(* IEC 61131-3 sources: daoli-st-library/DL_Process (part 17) *)

(* ---- FC_DL_RoRecoveryCalc.st ---- *)
(*
  Name: FC_DL_RoRecoveryCalc
  Category: DL_Process
  Version: 1.0.0
  Round: R90 / 2026-11-25
  开源溯源：clean-room 自研（族 RO/NF 膜法水处理，ST 开源生态实测 0 命中，无外部代码引入）
  功能：1) 系统回收率按「产水占进水的百分比」计算，产水为分子、进水为分母，方向固定不可交换，
           即 fRecoveryPct = fPermeateFlowM3h / fFeedFlowM3h * 100，用于 RO/NF 段回收率监视。
        2) 浓水排放流量由容积守恒的减法式给出：进水 − 产水（同温同压下的容积近似），
           作为浓水调节阀的前馈目标值使用。
        3) 回收率同时受两个独立门限约束：物理域 0.0 ~ 100.0 %，以及设计上限
           fRecoveryMaxPct（膜厂家给定的段回收率上限）；任一越界只置 xValid=FALSE，
           数值本身钳制到物理域内后输出，绝不把越限值伪装成合格值。
  边界条件：1) 分母零闸：ABS(fFeedFlowM3h) > DL_EPS 才允许做除法，否则清零全部输出并置无效。
        2) 非有限值闸：全部实值入参先过 NOT(x > -DL_BIG AND x < DL_BIG)，该式同时拦 NaN 与 Inf，
           命中即拦断实值通路（输出强制 0.0），不得只置标志而把 NaN 传给下游（R19）。
        3) 回收率物理域 0.0 ~ 100.0 %，越域钳制到域内输出并置 xValid=FALSE。
        4) 设计上限 fRecoveryMaxPct 自身须落在 (0.0, 100.0] 内，越域视为组态错误判无效。
        5) 产水量为负值（传感器反向）或大于进水量（超出守恒），均判无效，不取绝对值掩盖故障。
        6) 无回差环节：本件为纯函数无状态，不做迟滞，迟滞由下游报警件承担。
  量纲自证：fRecoveryPct = (m3/h) / (m3/h) * 100 = 无因次百分数 [%]；
           fBrineFlowM3h = (m3/h) − (m3/h) = (m3/h)，减法两侧同量纲，量纲关系合法。
*)

FUNCTION FC_DL_RoRecoveryCalc : BOOL
VAR_INPUT
    fFeedFlowM3h     : REAL;   // 系统进水体积流量 [m3/h] / Feed volumetric flow [m3/h]
    fPermeateFlowM3h : REAL;   // 系统产水体积流量 [m3/h] / Permeate volumetric flow [m3/h]
    fRecoveryMaxPct  : REAL;   // 段回收率设计上限 [%] / Design recovery upper limit [%]
END_VAR
VAR_OUTPUT
    fRecoveryPct     : REAL;   // 系统回收率 [%] / System recovery ratio [%]
    fBrineFlowM3h    : REAL;   // 浓水排放流量 [m3/h] / Brine discharge flow [m3/h]
    xValid           : BOOL;   // 计算有效标志 [bool] / Calculation valid flag [bool]
END_VAR
VAR
    _fRecRawPct      : REAL;   // 钳制前的原始回收率 [%] / Raw recovery before limiting [%]
    _fBrineRawM3h    : REAL;   // 钳制前的原始浓水流量 [m3/h] / Raw brine flow before limiting [m3/h]
END_VAR
VAR CONSTANT
    DL_EPS           : REAL := 1.0E-9;    // 分母零闸阈值 [-] / Division-zero gate threshold [-]
    DL_BIG           : REAL := 1.0E12;    // 非有限值闸量级上限 [-] / Finiteness gate magnitude [-]
    DL_PCT           : REAL := 100.0;     // 百分比换算因子 [%] / Percent conversion factor [%]
    DL_REC_LO_PCT    : REAL := 0.0;       // 回收率物理域下限 [%] / Recovery physical domain low [%]
    DL_REC_HI_PCT    : REAL := 100.0;     // 回收率物理域上限 [%] / Recovery physical domain high [%]
END_VAR

(* —— 段 1：非有限值闸（R19：闸断实值通路，NaN/Inf 一律不得流到输出） —— *)
IF NOT (fFeedFlowM3h > -DL_BIG AND fFeedFlowM3h < DL_BIG)
   OR NOT (fPermeateFlowM3h > -DL_BIG AND fPermeateFlowM3h < DL_BIG)
   OR NOT (fRecoveryMaxPct > -DL_BIG AND fRecoveryMaxPct < DL_BIG) THEN
    fRecoveryPct := 0.0;                    // 输出强制 0.0，切断污染源 / Force zero, cut polluted path
    fBrineFlowM3h := 0.0;                   // 浓水同样强制 0.0 / Brine forced to zero as well
    xValid := FALSE;                        // 有效位清零 / Validity cleared
    FC_DL_RoRecoveryCalc := FALSE;          // 返回码与有效位同源 / Return mirrors validity
    RETURN;                                 // 立即退出 / Immediate exit
END_IF

(* —— 段 2：分母零闸（R4：除法前先过 ABS 闸，且闸的是分母本身） —— *)
IF ABS(fFeedFlowM3h) <= DL_EPS THEN
    fRecoveryPct := 0.0;                    // 无进水即无回收率 / No feed means no recovery
    fBrineFlowM3h := 0.0;                   // 无进水即无浓水 / No feed means no brine
    xValid := FALSE;                        // 判无效 / Invalid
    FC_DL_RoRecoveryCalc := FALSE;          // 返回码同步 / Return synchronised
    RETURN;                                 // 提前退出，不做无意义运算 / Early exit
END_IF

(* —— 段 3：主算式（R22 方向自核：差值/比值的基准量是进水量，不是产水量） —— *)
_fRecRawPct := fPermeateFlowM3h / fFeedFlowM3h * DL_PCT;   // 产水 / 进水 * 100 [%]
_fBrineRawM3h := fFeedFlowM3h - fPermeateFlowM3h;          // 进水 − 产水 [m3/h]

(* —— 段 4：物理域与设计上限校验（单点 BOOL 聚合，避免多处赋 FALSE 造成覆盖） —— *)
xValid := (_fRecRawPct >= DL_REC_LO_PCT)                       // 不低于物理域下限
          AND (_fRecRawPct <= DL_REC_HI_PCT)                   // 不高于物理域上限
          AND (fRecoveryMaxPct > DL_EPS)                       // 设计上限必须为正
          AND (fRecoveryMaxPct <= DL_REC_HI_PCT)               // 设计上限不得超 100 %
          AND (_fRecRawPct <= fRecoveryMaxPct)                 // 不得超出膜厂家设计上限
          AND (fPermeateFlowM3h >= 0.0)                        // 产水不得为负（传感器反向）
          AND (fPermeateFlowM3h <= fFeedFlowM3h)               // 产水不得大于进水（守恒校验）
          AND (_fBrineRawM3h >= 0.0);                          // 浓水不得为负

(* —— 段 5：输出单点写盘（数值钳制到物理域内，有效位已在段 4 定案） —— *)
fRecoveryPct := LIMIT(DL_REC_LO_PCT, _fRecRawPct, DL_REC_HI_PCT);   // 回收率钳 0..100 [%]
fBrineFlowM3h := MAX(DL_REC_LO_PCT, _fBrineRawM3h);                 // 浓水钳 >= 0 [m3/h]
FC_DL_RoRecoveryCalc := xValid;                                     // 返回码：TRUE = 计算可信

END_FUNCTION

(* ---- FC_DL_RoScaleSaturationIndexCalc.st ---- *)
(*
  Name: FC_DL_RoScaleSaturationIndexCalc
  Category: DL_Process
  Version: 1.0.0
  Round: R90 / 2026-11-25
  开源溯源：clean-room 自研（族 RO/NF 膜法水处理，ST 开源生态实测 0 命中，无外部代码引入）
  功能：1) 朗格利尔饱和指数按经典四因子式解算：LSI = pH − pHs，
           其中 pHs = (9.3 + A + B) − (C + D)：
             A = (LOG10(TDS) − 1) / 10，表征溶解固体的离子强度；
             B = −13.12 · LOG10(T_K) + 34.55，温度项（T_K 为开尔文，必须做 °C→K 偏移）；
             C = LOG10(Ca 硬度) − 0.4，钙硬度项；
             D = LOG10(碱度)，碱度项。
        2) LOG10 用跨平台安全写法 LN(x) / LN(10) 实现，不依赖厂商私有 LOG10 扩展。
        3) 输出结垢风险等级整数 iRiskLvl：0 = 不结垢（偏腐蚀），1 = 轻度结垢，
           2 = 中度结垢，3 = 严重结垢；等级由 LSI 阈值判定，供加药/阻垢剂投加策略直接取用。
  边界条件：1) 非有限值闸：五路实值入参统一过 NOT(x > -DL_BIG AND x < DL_BIG)，
           同时拦 NaN 与 Inf，命中即拦断实值通路（fLsi 强制 0.0、iRiskLvl 置 0）并置无效（R19）。
        2) 对数自变量零闸：TDS / 钙硬度 / 碱度三项都必须 ABS(x) > DL_EPS 才可进 LN，
           否则 LOG10 发散；任一项不满足判无效。
        3) 对数自变量负值闸：三量均为浓度，负值属变送器故障，判无效且不取 ABS 掩盖。
        4) 量程钳制：TDS 钳 0..60000 mg/L、钙硬度与碱度钳 0..DL_HARD_MAX(2000 mg/L)、
           pH 钳 0..14、温度钳 0..90 °C；越域钳边界值参与计算但置无效。
        5) LSI 结果饱和钳到 −5.0 ~ +5.0 的工程可观测域，防极端输入把指数推到无意义量级。
        6) 无回差环节：纯函数无状态，等级切换的迟滞由下游报警件承担。
  量纲自证：A = (LOG10(mg/L) − 1) / 10 → 无因次 [-]，LOG10 的自变量已按 mg/L 归一；
           B = −13.12 · LOG10(K) + 34.55 → 无因次 [-]，34.55 为经验截距，无单位；
           C、D 同 A 均为无因次；LSI = pH(−) − pHs(−) = 无因次指数 [-]，四项量纲一致。
*)

FUNCTION FC_DL_RoScaleSaturationIndexCalc : BOOL
VAR_INPUT
    fPh              : REAL;   // 给水 pH 值 [pH 单位] / Feed water pH [pH unit]
    fTempC           : REAL;   // 给水温度 [°C] / Feed water temperature [°C]
    fCaHardnessMgL   : REAL;   // 钙硬度（以 CaCO3 计）[mg/L] / Calcium hardness as CaCO3 [mg/L]
    fAlkalinityMgL   : REAL;   // 总碱度（以 CaCO3 计）[mg/L] / Total alkalinity as CaCO3 [mg/L]
    fTdsMgL          : REAL;   // 总溶解固体 [mg/L] / Total dissolved solids [mg/L]
END_VAR
VAR_OUTPUT
    fLsi             : REAL;   // 朗格利尔饱和指数 [-] / Langelier saturation index [-]
    iRiskLvl         : INT;    // 结垢风险等级 0..3 [-] / Scaling risk level 0..3 [-]
    xValid           : BOOL;   // 计算有效标志 [bool] / Calculation valid flag [bool]
END_VAR
VAR
    _fPhClamp        : REAL;   // 钳制后的 pH [-] / Clamped pH [-]
    _fTClampC        : REAL;   // 钳制后的温度 [°C] / Clamped temperature [°C]
    _fCaClampMgL     : REAL;   // 钳制后的钙硬度 [mg/L] / Clamped calcium hardness [mg/L]
    _fAlkClampMgL    : REAL;   // 钳制后的碱度 [mg/L] / Clamped alkalinity [mg/L]
    _fTdsClampMgL    : REAL;   // 钳制后的 TDS [mg/L] / Clamped TDS [mg/L]
    _fTermA          : REAL;   // A 项（TDS 项）[-] / Term A, TDS term [-]
    _fTermB          : REAL;   // B 项（温度项）[-] / Term B, temperature term [-]
    _fTermC          : REAL;   // C 项（钙硬度项）[-] / Term C, calcium hardness term [-]
    _fTermD          : REAL;   // D 项（碱度项）[-] / Term D, alkalinity term [-]
    _fPhs            : REAL;   // 饱和 pH [-] / Saturation pH [-]
    _fLsiRaw         : REAL;   // 未饱和的原始 LSI [-] / Raw LSI before limiting [-]
    _bLogOk          : BOOL;   // 对数自变量合法性聚合 [-] / Logarithm argument validity aggregate
END_VAR
VAR CONSTANT
    DL_EPS           : REAL := 1.0E-9;    // 对数自变量零闸阈值 [-] / Logarithm argument zero gate [-]
    DL_BIG           : REAL := 1.0E12;    // 非有限值闸量级上限 [-] / Finiteness gate magnitude [-]
    DL_K0            : REAL := 273.15;    // 摄氏转开尔文偏移 [K] / Celsius to Kelvin offset [K]
    DL_LN10          : REAL := 2.302585093;   // LN(10)，用于实现 LOG10 [-] / LN(10) for LOG10 [-]
    DL_PH_MAX        : REAL := 14.0;      // pH 量程上限 [-] / pH range high [-]
    DL_T_HI_C        : REAL := 90.0;      // 温度量程上限 [°C] / Temperature range high [°C]
    DL_HARD_MAX      : REAL := 2000.0;    // 钙硬度/碱度量程上限 [mg/L] / Hardness range high [mg/L]
    DL_TDS_MAX       : REAL := 60000.0;   // TDS 量程上限 [mg/L] / TDS range high [mg/L]
    DL_LSI_LO        : REAL := -5.0;      // LSI 工程可观测下限 [-] / LSI observable low [-]
    DL_LSI_HI        : REAL := 5.0;       // LSI 工程可观测上限 [-] / LSI observable high [-]
    DL_LSI_L1        : REAL := 0.0;       // 等级 0/1 分界 [-] / Risk level 0-to-1 boundary [-]
    DL_LSI_L2        : REAL := 0.5;       // 等级 1/2 分界 [-] / Risk level 1-to-2 boundary [-]
    DL_LSI_L3        : REAL := 1.5;       // 等级 2/3 分界 [-] / Risk level 2-to-3 boundary [-]
END_VAR

(* —— 段 1：非有限值闸（R19：五路入参全覆盖，拦 NaN 与 Inf） —— *)
IF NOT (fPh > -DL_BIG AND fPh < DL_BIG)
   OR NOT (fTempC > -DL_BIG AND fTempC < DL_BIG)
   OR NOT (fCaHardnessMgL > -DL_BIG AND fCaHardnessMgL < DL_BIG)
   OR NOT (fAlkalinityMgL > -DL_BIG AND fAlkalinityMgL < DL_BIG)
   OR NOT (fTdsMgL > -DL_BIG AND fTdsMgL < DL_BIG) THEN
    fLsi := 0.0;                            // 输出强制 0.0 / Output forced to zero
    iRiskLvl := 0;                          // 等级置 0（不结垢），不给误导性等级 / Risk level cleared
    xValid := FALSE;                        // 有效位清零 / Validity cleared
    FC_DL_RoScaleSaturationIndexCalc := FALSE;   // 返回码同源 / Return mirrors validity
    RETURN;                                 // 立即退出 / Immediate exit
END_IF

(* —— 段 2：对数自变量零闸 + 负值闸（R4：LN 的自变量必须先验正） —— *)
_bLogOk := (fTdsMgL > DL_EPS) AND (fCaHardnessMgL > DL_EPS) AND (fAlkalinityMgL > DL_EPS);
IF NOT _bLogOk THEN
    fLsi := 0.0;                            // 输出强制 0.0 / Output forced to zero
    iRiskLvl := 0;                          // 等级置 0 / Risk level cleared
    xValid := FALSE;                        // 判无效 / Invalid
    FC_DL_RoScaleSaturationIndexCalc := FALSE;   // 返回码同步 / Return synchronised
    RETURN;                                 // 提前退出 / Early exit
END_IF

(* —— 段 3：量程钳制（边界值参与计算，越域在段 5 判无效） —— *)
_fPhClamp := LIMIT(0.0, fPh, DL_PH_MAX);                  // pH 钳 0..14 [-]
_fTClampC := LIMIT(0.0, fTempC, DL_T_HI_C);               // 温度钳 0..90 [°C]
_fCaClampMgL := LIMIT(0.0, fCaHardnessMgL, DL_HARD_MAX);  // 钙硬度钳 [mg/L]
_fAlkClampMgL := LIMIT(0.0, fAlkalinityMgL, DL_HARD_MAX); // 碱度钳 [mg/L]
_fTdsClampMgL := LIMIT(0.0, fTdsMgL, DL_TDS_MAX);         // TDS 钳 [mg/L]

(* —— 段 4：四因子解算（LOG10 以 LN(x)/LN(10) 跨平台实现） —— *)
_fTermA := (LN(_fTdsClampMgL) / DL_LN10 - 1.0) / 10.0;                          // A 项 [-]
_fTermB := -13.12 * (LN(_fTClampC + DL_K0) / DL_LN10) + 34.55;                  // B 项 [-]
_fTermC := LN(_fCaClampMgL) / DL_LN10 - 0.4;                                    // C 项 [-]
_fTermD := LN(_fAlkClampMgL) / DL_LN10;                                         // D 项 [-]
_fPhs := (9.3 + _fTermA + _fTermB) - (_fTermC + _fTermD);                       // 饱和 pH [-]
_fLsiRaw := _fPhClamp - _fPhs;                                                  // LSI = pH − pHs [-]

(* —— 段 5：有效位单点聚合（量程校验，钳制值已参与计算） —— *)
xValid := (fPh >= 0.0) AND (fPh <= DL_PH_MAX)                                   // pH 在量程内
          AND (fTempC >= 0.0) AND (fTempC <= DL_T_HI_C)                         // 温度在量程内
          AND (fCaHardnessMgL <= DL_HARD_MAX)                                   // 钙硬度不越上限
          AND (fAlkalinityMgL <= DL_HARD_MAX)                                   // 碱度不越上限
          AND (fTdsMgL <= DL_TDS_MAX);                                          // TDS 不越上限

(* —— 段 6：风险等级分级（IF/ELSIF 单链，iRiskLvl 只在此处赋值一次） —— *)
IF _fLsiRaw < DL_LSI_L1 THEN
    iRiskLvl := 0;                          // 不结垢（偏腐蚀倾向）/ Non-scaling, corrosive tendency
ELSIF _fLsiRaw < DL_LSI_L2 THEN
    iRiskLvl := 1;                          // 轻度结垢 / Slight scaling tendency
ELSIF _fLsiRaw < DL_LSI_L3 THEN
    iRiskLvl := 2;                          // 中度结垢 / Moderate scaling tendency
ELSE
    iRiskLvl := 3;                          // 严重结垢 / Severe scaling tendency
END_IF

(* —— 段 7：输出单点写盘（LSI 饱和钳到工程可观测域） —— *)
fLsi := LIMIT(DL_LSI_LO, _fLsiRaw, DL_LSI_HI);   // LSI 钳 −5..+5 [-]
FC_DL_RoScaleSaturationIndexCalc := xValid;      // 返回码：TRUE = 计算可信

END_FUNCTION

(* ---- FC_DL_RoStagePressureDropCalc.st ---- *)
(*
  Name: FC_DL_RoStagePressureDropCalc
  Category: DL_Process
  Version: 1.0.0
  Round: R90 / 2026-11-25
  开源溯源：clean-room 自研（族 RO/NF 膜法水处理，ST 开源生态实测 0 命中，无外部代码引入）
  功能：1) 段间压降按湍流平方律计算：ΔP = k · Q²，其中 k 为段阻力系数（bar/(m3/h)²），
           Q 为段流量（m3/h）。平方律的依据是湍流区沿程与局部损失均与流速平方成正比，
           而流速与容积流量成正比，故压降对流量呈二次关系，不是线性关系。
        2) 与压降上限 fDropLimitBar 比对给出超限报警 xAlarm。超限是膜段污堵/浓水通道阻塞的
           早期特征（流量不变而压降上升），因此报警取「大于等于上限」而非「大于」，
           上限触点本身即算到达报警点。
  边界条件：1) 非有限值闸：三路实值入参统一过 NOT(x > -DL_BIG AND x < DL_BIG)，
           同时拦 NaN 与 Inf，命中即拦断实值通路（fDropBar 强制 0.0、xAlarm 强制 FALSE）并置无效（R19）。
        2) 组态零闸：ABS(fResistCoef) > DL_EPS 与 ABS(fDropLimitBar) > DL_EPS 都必须成立，
           阻力系数为 0 表示未标定、上限为 0 表示未组态，两者都判无效（不做除零以外的默认替代）。
        3) 负值闸：段流量为负判无效（传感器反向）；阻力系数为负判无效（系数不可为负）；
           压降上限为负判无效。
        4) 饱和钳制：段流量先钳到 0 ~ DL_FLOW_MAX(1000 m3/h)，压降结果再钳到 0 ~ DL_DROP_MAX(50 bar)，
           防止平方项在小数域溢出或给出无物理意义的巨值。
        5) 报警只在 xValid 为 TRUE 时才可能为 TRUE，无效数据不得触发工艺报警（防误停）。
        6) 无回差环节：本件为纯函数无状态，报警回差由下游 FB 承担。
  量纲自证：ΔP = (bar/(m3/h)²) × (m3/h)² = bar，平方项与系数分母量纲对消，量纲闭合；
           报警比较两侧同为 bar，量纲一致，禁止与 kPa 混比。
*)

FUNCTION FC_DL_RoStagePressureDropCalc : BOOL
VAR_INPUT
    fStageFlowM3h    : REAL;   // 段内体积流量 [m3/h] / Stage volumetric flow [m3/h]
    fResistCoef      : REAL;   // 段阻力系数 [bar/(m3/h)²] / Stage resistance coefficient [bar/(m3/h)^2]
    fDropLimitBar    : REAL;   // 段间压降报警上限 [bar] / Pressure drop alarm limit [bar]
END_VAR
VAR_OUTPUT
    fDropBar         : REAL;   // 段间压降 [bar] / Stage pressure drop [bar]
    xAlarm           : BOOL;   // 压降超限报警 [bool] / Pressure drop over-limit alarm [bool]
    xValid           : BOOL;   // 计算有效标志 [bool] / Calculation valid flag [bool]
END_VAR
VAR
    _fFlowClampM3h   : REAL;   // 钳制后的段流量 [m3/h] / Clamped stage flow [m3/h]
    _fDropRawBar     : REAL;   // 未饱和的原始压降 [bar] / Raw pressure drop [bar]
END_VAR
VAR CONSTANT
    DL_EPS           : REAL := 1.0E-9;    // 组态零闸阈值 [-] / Configuration zero gate threshold [-]
    DL_BIG           : REAL := 1.0E12;    // 非有限值闸量级上限 [-] / Finiteness gate magnitude [-]
    DL_FLOW_MAX      : REAL := 1000.0;    // 段流量饱和钳制上限 [m3/h] / Stage flow saturation ceiling [m3/h]
    DL_DROP_MAX      : REAL := 50.0;      // 压降饱和钳制上限 [bar] / Pressure drop saturation ceiling [bar]
END_VAR

(* —— 段 1：非有限值闸（R19：三路入参全覆盖，拦 NaN 与 Inf） —— *)
IF NOT (fStageFlowM3h > -DL_BIG AND fStageFlowM3h < DL_BIG)
   OR NOT (fResistCoef > -DL_BIG AND fResistCoef < DL_BIG)
   OR NOT (fDropLimitBar > -DL_BIG AND fDropLimitBar < DL_BIG) THEN
    fDropBar := 0.0;                        // 输出强制 0.0 / Output forced to zero
    xAlarm := FALSE;                        // 报警强制 FALSE，无效数据不得触发停运 / Alarm forced off
    xValid := FALSE;                        // 有效位清零 / Validity cleared
    FC_DL_RoStagePressureDropCalc := FALSE; // 返回码同源 / Return mirrors validity
    RETURN;                                 // 立即退出 / Immediate exit
END_IF

(* —— 段 2：组态零闸（阻力系数与报警上限都必须已标定，0 值视为未组态） —— *)
IF (ABS(fResistCoef) <= DL_EPS) OR (ABS(fDropLimitBar) <= DL_EPS) THEN
    fDropBar := 0.0;                        // 输出强制 0.0 / Output forced to zero
    xAlarm := FALSE;                        // 报警强制 FALSE / Alarm forced off
    xValid := FALSE;                        // 判无效 / Invalid
    FC_DL_RoStagePressureDropCalc := FALSE; // 返回码同步 / Return synchronised
    RETURN;                                 // 提前退出 / Early exit
END_IF

(* —— 段 3：负值闸（流量反向 / 系数为负 / 上限为负，三者均属组态或传感器故障） —— *)
IF (fStageFlowM3h < 0.0) OR (fResistCoef < 0.0) OR (fDropLimitBar < 0.0) THEN
    fDropBar := 0.0;                        // 输出强制 0.0 / Output forced to zero
    xAlarm := FALSE;                        // 报警强制 FALSE / Alarm forced off
    xValid := FALSE;                        // 判无效 / Invalid
    FC_DL_RoStagePressureDropCalc := FALSE; // 返回码同步 / Return synchronised
    RETURN;                                 // 提前退出 / Early exit
END_IF

(* —— 段 4：平方律主算式（R22 方向自核：流量平方乘系数，非系数除流量） —— *)
_fFlowClampM3h := LIMIT(0.0, fStageFlowM3h, DL_FLOW_MAX);    // 流量钳 0..1000 [m3/h]
_fDropRawBar := fResistCoef * _fFlowClampM3h * _fFlowClampM3h;   // ΔP = k·Q² [bar]

(* —— 段 5：输出单点写盘（先饱和钳制，再据此判报警，保证判据用的是同一个值） —— *)
fDropBar := LIMIT(0.0, _fDropRawBar, DL_DROP_MAX);           // 压降钳 0..50 [bar]
xValid := (fResistCoef > DL_EPS)                             // 系数已标定且为正
          AND (fDropLimitBar > DL_EPS)                       // 上限已组态且为正
          AND (fStageFlowM3h >= 0.0);                        // 流量非负
xAlarm := xValid AND (fDropBar >= fDropLimitBar);            // 到达上限即报警（含触点）

(* —— 段 6：返回码（TRUE = 计算可信，与 xValid 同源） —— *)
FC_DL_RoStagePressureDropCalc := xValid;

END_FUNCTION

(* ---- FC_DL_SandToMetalRatioCalc.st ---- *)
(*
 * FC_DL_SandToMetalRatioCalc | C1 | DL_Process
 * 功能：砂铁比（单位铸铁合格件对应的砂循环量）       单位：流量 [kg/h]、比值 [kg/kg]
 * 工况边界：仅适用于连续生产的砂处理线（砂循环量与铁水消耗量同口径统计）；金属流量须 >0（入分母），砂流量须 ≥0 且有限；不区分新旧砂，只算总量比值
 * 代数值回代：sand=120000 kg/h、metal=15000 kg/h → 比值 8.0 kg/kg（与 spec 回代行一致）
 * 开源溯源：clean-room 自研，未复制任何第三方代码（无外部来源）
 *)
FUNCTION FC_DL_SandToMetalRatioCalc : BOOL
VAR_INPUT
    rSandKgH  : REAL := 120000.0;    // 砂循环量 | sand circulation rate [kg/h]
    rMetalKgH : REAL := 15000.0;     // 铁水消耗量 | molten metal consumption rate [kg/h]
END_VAR
VAR_OUTPUT
    rRatio     : REAL;               // 砂铁比 | sand to metal ratio [kg/kg]
    xValid     : BOOL;               // 输出有效 | outputs valid
    nFaultCode : INT;                // 0=无 / 9711=金属流量非法 | 0 none, 9711 illegal metal flow
END_VAR
VAR
    xFinSand  : BOOL;                // 砂流量有限性 | sand flow is finite
    xFinMetal : BOOL;                // 金属流量有限性 | metal flow is finite
END_VAR
VAR CONSTANT
    DL_SMR_METAL_MIN : REAL := 1.0E-9;  // 金属流量下限（防零除）| metal flow lower bound [kg/h]
END_VAR

// 段1｜非有限闸（R19）
xFinSand := (rSandKgH = rSandKgH) AND ((rSandKgH - rSandKgH) = 0.0);
xFinMetal := (rMetalKgH = rMetalKgH) AND ((rMetalKgH - rMetalKgH) = 0.0);
IF (NOT xFinSand) OR (NOT xFinMetal) THEN
    rRatio := 0.0;                   // 安全值：比值 0 | safe value, zero ratio
    xValid := FALSE;
    nFaultCode := 9711;
    FC_DL_SandToMetalRatioCalc := FALSE;
    RETURN;
END_IF

// 段2｜域闸：金属流量入分母必须 >0，砂流量不得为负
IF (rMetalKgH <= DL_SMR_METAL_MIN) OR (rSandKgH < 0.0) THEN
    rRatio := 0.0;
    xValid := FALSE;
    nFaultCode := 9711;
    FC_DL_SandToMetalRatioCalc := FALSE;
    RETURN;
END_IF

// 段3｜算法与出口
rRatio := rSandKgH / rMetalKgH;
nFaultCode := 0;
xValid := TRUE;
FC_DL_SandToMetalRatioCalc := TRUE;
END_FUNCTION

(* ---- FC_DL_SanitizeHoldTimeCalc.st ---- *)
(*
  ============================================================
  组件名 : FC_DL_SanitizeHoldTimeCalc
  分类   : DL_Process
  功能   : 消毒保持时间计算，按实际浓度折算浓度比并对温度系数修正后给出保持时间
  复杂度 : C1
  版本   : 1.0.0
  作者   : 道莅工业代码库工厂 / R81
  日期   : 2026-11-24
  开源溯源 : clean-room（no upstream）—— 依据公开工程公式自研，未复制任何上游实现
  红线自检 : R1 无GVL/R2 无物理地址/R3 纯IEC/R4 防除零/R5 双语注释
  接口说明 :
      温度系数 = 1 + (温度-20)*0.02，限幅 0.5~2.0，防止极端温度把时间推到无意义区间。
      保持时间 = 基准时间 * (基准浓度/实际浓度) * (1/温度系数)。
      浓度低于基准时比值大于 1，时间自动延长；浓度高于基准时时间缩短，符合消毒动力学方向。
  ============================================================
*)
FUNCTION FC_DL_SanitizeHoldTimeCalc : BOOL
VAR_INPUT
    bEnable      : BOOL; // 使能：TRUE 时计算 / Enable: TRUE to compute
    bErr         : BOOL; // 外部故障：TRUE 时立即退出并置结果无效 / External fault: TRUE aborts with invalid result
    rConcPct     : REAL; // 实际消毒液浓度 [%] / actual sanitizer concentration [percent]
    rConcRefPct  : REAL; // 基准消毒液浓度 [%] / reference sanitizer concentration [percent]
    rHoldRef_min : REAL; // 基准浓度下的基准保持时间 [min] / reference hold time at the reference concentration [minute]
    rTempC       : REAL; // 实际消毒液温度 [摄氏度] / actual sanitizer temperature [degree Celsius]
END_VAR
VAR_OUTPUT
    rTempFactor : REAL; // 温度修正系数，限幅 0.5~2.0 [无量纲] / temperature correction factor clamped to 0.5 to 2.0 [dimensionless]
    rConcRatio  : REAL; // 浓度比，基准浓度除以实际浓度 [无量纲] / concentration ratio of reference over actual [dimensionless]
    rHold_min   : REAL; // 修正后的保持时间 [min] / corrected hold time [minute]
    bValid      : BOOL; // 输出有效：TRUE 表示结果可用 / Output valid
END_VAR
VAR CONSTANT
    DL_R_MAX    : REAL := 3.0E38; // 实数上界，用于拦截 Inf [无量纲] / real upper bound used to reject infinity [dimensionless]
    DL_EPS      : REAL := 1.0E-12; // 除零判定阈值 [无量纲] / division guard threshold [dimensionless]
    DL_ONE      : REAL := 1.0;    // 单位常量 [无量纲] / unity constant [dimensionless]
    DL_TEMP_REF : REAL := 20.0;   // 温度基准点 [摄氏度] / temperature reference point [degree Celsius]
    DL_TEMP_K   : REAL := 0.02;   // 每摄氏度温度系数增量 [1/摄氏度] / temperature coefficient increment per degree Celsius [per degree Celsius]
    DL_FACT_LO  : REAL := 0.5;    // 温度系数下限 [无量纲] / lower limit of the temperature factor [dimensionless]
    DL_FACT_HI  : REAL := 2.0;    // 温度系数上限 [无量纲] / upper limit of the temperature factor [dimensionless]
    DL_TEMP_MIN : REAL := -50.0;  // 允许温度下界 [摄氏度] / permitted lower bound of the temperature [degree Celsius]
    DL_TEMP_MAX : REAL := 150.0;  // 允许温度上界 [摄氏度] / permitted upper bound of the temperature [degree Celsius]
END_VAR
VAR
    _bFin  : BOOL := FALSE; // 输入有限性判定结果 / input finiteness verdict
    _rInv  : REAL := 0.0;   // 温度系数的倒数，除法前先算后判 [无量纲] / reciprocal of the temperature factor computed before the guard [dimensionless]
END_VAR

    // 段 1｜出口预置：系数先置于 1，避免下游误用零
    rTempFactor := DL_ONE;
    rConcRatio := 0.0;
    rHold_min := 0.0;
    bValid := FALSE;
    // 段 2｜使能闸与外部故障闸
    IF NOT bEnable THEN
        RETURN;
    END_IF;
    IF bErr THEN
        RETURN;
    END_IF;
    // 段 3｜非有限闸
    _bFin := (rConcPct = rConcPct) AND (ABS(rConcPct) <= DL_R_MAX) AND (rConcRefPct = rConcRefPct) AND (ABS(rConcRefPct) <= DL_R_MAX) AND (rHoldRef_min = rHoldRef_min) AND (ABS(rHoldRef_min) <= DL_R_MAX) AND (rTempC = rTempC) AND (ABS(rTempC) <= DL_R_MAX);
    IF NOT _bFin THEN
        RETURN;
    END_IF;
    // 段 4｜域闸：实际浓度严格为正、基准浓度非负、基准时间非负、温度在工程区间
    IF ABS(rConcPct) <= DL_EPS THEN
        RETURN;
    END_IF;
    IF (rConcPct < 0.0) OR (rConcRefPct < 0.0) OR (rHoldRef_min < 0.0) THEN
        RETURN;
    END_IF;
    IF (rTempC < DL_TEMP_MIN) OR (rTempC > DL_TEMP_MAX) THEN
        RETURN;
    END_IF;
    // 段 5｜温度系数与限幅
    rTempFactor := DL_ONE + (rTempC - DL_TEMP_REF) * DL_TEMP_K;
    IF rTempFactor > DL_FACT_HI THEN
        rTempFactor := DL_FACT_HI;
    ELSIF rTempFactor < DL_FACT_LO THEN
        rTempFactor := DL_FACT_LO;
    END_IF;
    // 段 6｜浓度比
    rConcRatio := rConcRefPct / rConcPct;
    // 段 7｜温度系数分母闸：先判零再取倒数，顺序不可颠倒
    IF ABS(rTempFactor) <= DL_EPS THEN
        RETURN;
    END_IF;
    _rInv := DL_ONE / rTempFactor;
    rHold_min := rHoldRef_min * rConcRatio * _rInv;
    bValid := TRUE;
    FC_DL_SanitizeHoldTimeCalc := bValid;
END_FUNCTION

(* ---- FC_DL_ScreenEfficiencyCalc.st ---- *)
(*
  Name: FC_DL_ScreenEfficiencyCalc
  Category: DL_Process
  Version: 1.0.0
  Round: R89 / 2026-11-25
  开源溯源：clean-room 自研（族 矿山破碎筛分，ST 开源生态实测 0 命中，无外部代码引入）
  功能：按入料/筛上/筛下三处细粒含量算振动筛筛分效率（经典式，全部折算为小数参与运算）。
  边界条件：① 三入参百分数先折算小数，入料细粒 0~100 %、筛上 0~100 %、筛下 0~100 %；
            ② 分母 (1−O)·(F+U−1) 显式零闸，绝对值不超 DL_EPS 即判非法返回哨兵 -1；
            ③ 效率物理域 0~100 %；算得负值（物料衡算矛盾，如筛下含量低于入料）判 xValid = FALSE 并返回 -1。
  量纲自证：F/O/U 均为质量分数（无量纲），E 亦无量纲，×100 得百分数。
*)
FUNCTION FC_DL_ScreenEfficiencyCalc : REAL
VAR_INPUT
    fFeedFinesPct : REAL;   (* 入料细粒含量 [%] Feed fines content [%] *)
    fOverFinesPct : REAL;   (* 筛上细粒含量 [%] Oversize fines content [%] *)
    fUnderFinesPct : REAL;  (* 筛下合格细粒含量 [%] Undersize fines content [%] *)
END_VAR
VAR_OUTPUT
    fEfficiencyPct : REAL;  (* 筛分效率 [%] Screening efficiency [%] *)
    xValid : BOOL;          (* 计算有效性标志 [-] Calculation valid flag *)
END_VAR
VAR CONSTANT
    DL_EPS : REAL := 1.0E-9;    (* 除零判定容差 [-] Divide-by-zero tolerance *)
    DL_PCT : REAL := 100.0;     (* 百分数基准 [%] Percent base *)
    DL_E_MAX : REAL := 100.0;   (* 效率饱和上限 [%] Efficiency ceiling *)
END_VAR
VAR
    fF : REAL;      (* 入料细粒质量分数 [-] Feed fines fraction *)
    fO : REAL;      (* 筛上细粒质量分数 [-] Oversize fines fraction *)
    fU : REAL;      (* 筛下细粒质量分数 [-] Undersize fines fraction *)
    fDen : REAL;    (* 分母 (1−O)·(F+U−1) [-] Denominator *)
    fEff : REAL;    (* 效率小数中间量 [-] Efficiency scratch *)
END_VAR
(* 出口预置：两出口统一预置（R256） *)
fEfficiencyPct := 0.0; xValid := FALSE;
(* 非有限闸：NaN 自反判 + Inf 差值自减判，三入参全枚举 *)
IF (fFeedFinesPct <> fFeedFinesPct) OR ((fFeedFinesPct - fFeedFinesPct) <> 0.0)
   OR (fOverFinesPct <> fOverFinesPct) OR ((fOverFinesPct - fOverFinesPct) <> 0.0)
   OR (fUnderFinesPct <> fUnderFinesPct) OR ((fUnderFinesPct - fUnderFinesPct) <> 0.0) THEN
    FC_DL_ScreenEfficiencyCalc := -1.0;     (* 哨兵 -1：入参非有限 / Sentinel -1, non-finite input *)
    RETURN;
END_IF
(* 组态域闸：三处含量皆须落在 0~100 %，入料细粒须 > 0（为除子） *)
IF (fFeedFinesPct <= DL_EPS) OR (fFeedFinesPct > DL_PCT)
   OR (fOverFinesPct < 0.0) OR (fOverFinesPct >= DL_PCT)
   OR (fUnderFinesPct < 0.0) OR (fUnderFinesPct > DL_PCT) THEN
    FC_DL_ScreenEfficiencyCalc := -1.0;     (* 哨兵 -1：组态非法 / Sentinel -1, bad configuration *)
    RETURN;
END_IF
(* 百分数折算小数，量纲变为质量分数 *)
fF := fFeedFinesPct / DL_PCT;
fO := fOverFinesPct / DL_PCT;
fU := fUnderFinesPct / DL_PCT;
(* 经典二产品筛分效率式分母：D = F·(U−O)，先算后闸，禁先除后判 *)
(* 原式 D=(1−O)(F+U−1) 会把 η 放大 1/(F+U−1) 倍并系统性饱和到 100%，已废弃 *)
fDen := fF * (fU - fO);
IF ABS(fDen) <= DL_EPS THEN
    FC_DL_ScreenEfficiencyCalc := -1.0;     (* 哨兵 -1：分母塌零 / Sentinel -1, vanishing denominator *)
    RETURN;
END_IF
(* E = U·(F−O) / (F·(U−O))，F 已过零闸，D 已过塌零闸（Wills 选矿手册式） *)
fEff := (fU * (fF - fO)) / fDen;
(* 负值即物料衡算矛盾（筛下细粒反少于入料平衡），判非法不钳成 0 冒充正常 *)
IF fEff < -DL_EPS THEN
    FC_DL_ScreenEfficiencyCalc := -1.0;     (* 哨兵 -1：衡算矛盾 / Sentinel -1, mass-balance conflict *)
    RETURN;
END_IF
(* 物理域钳位：效率不超 100 %，微负残差按 0 处理 *)
IF fEff > 1.0 THEN
    fEff := 1.0;                            (* 上限钳位 100 % / Clamp to 100 percent *)
ELSIF fEff < 0.0 THEN
    fEff := 0.0;                            (* 微负残差归零 / Negative residual to zero *)
END_IF
fEfficiencyPct := fEff * DL_PCT;            (* 分数 → 百分数 [%] Fraction to percent *)
xValid := TRUE;                             (* 链路有效 / Chain valid *)
FC_DL_ScreenEfficiencyCalc := fEfficiencyPct;
END_FUNCTION

(* ---- FC_DL_ScrewPressThroughput.st ---- *)
(*
  道莅工业代码库 / Daoli Industrial ST Library
  组件: FC_DL_ScrewPressThroughput
  分类: DL_Process
  开源溯源: 无（clean-room 工程公式自研；参考公开工艺计算公式，未复制任何受版权保护代码）
  许可证: 本项目自有 (MIT)
  功能: 螺旋压榨机干固体（DS）处理量换算：小时量与按日运行小时数折算的日总量
*)
FUNCTION FC_DL_ScrewPressThroughput : BOOL
VAR_INPUT
    rFlowM3h : REAL; // 进泥体积流量 [m3/h] / sludge feed flow
    rTsPct : REAL; // 进泥含固率 [%] / feed total solids content
    rRunHours : REAL; // 日运行小时数 [h/d] / daily running hours
END_VAR
VAR_OUTPUT
    rDsKgH : REAL; // 干固体小时处理量 [kg/h] / dry solids throughput per hour
    rDsKgDay : REAL; // 干固体日处理量 [kg/d] / dry solids throughput per day
    bValid : BOOL; // 结果有效位 [-] / result valid flag
    iErrCode : INT; // 事件码 0=正常 1=含固率超域 2=运行小时超域 3=结果非有限 / event code
END_VAR
VAR CONSTANT
    rRhoSludge : REAL := 1000.0; // 污泥近似密度 [kg/m3] / approximate sludge density
    rPctToFrac : REAL := 0.01; // 百分数转小数系数 [-]/[%] / percent to fraction factor
    rHourPerDay : REAL := 24.0; // 每日小时数 [h/d] / hours per day
END_VAR
VAR
    rDsRaw : REAL; // 未校验小时量 [kg/h] / unchecked hourly throughput
END_VAR

    // —— 段 0：全路径预清 —— //
    rDsRaw := 0.0;
    rDsKgH := 0.0;
    rDsKgDay := 0.0;
    bValid := FALSE;
    iErrCode := 0;
    FC_DL_ScrewPressThroughput := FALSE;
    // —— 段 1：含固率域闸 (0, 100]% —— //
    IF (rTsPct <= 0.0) OR (rTsPct > 100.0) THEN
        iErrCode := 1; // 含固率超域，干固体量无意义 / TS out of domain, dry solids meaningless
        RETURN;
    END_IF;
    // —— 段 2：日运行小时域闸 (0, 24]h —— //
    IF (rRunHours <= 0.0) OR (rRunHours > rHourPerDay) THEN
        iErrCode := 2; // 运行小时超域 / running hours out of domain
        RETURN;
    END_IF;
    // —— 段 3：量纲链 (m3/h)*(kg/m3)*(%)*(0.01) = kg/h —— //
    rDsRaw := rFlowM3h * rRhoSludge * rTsPct * rPctToFrac; // 干固体量 [kg/h] / dry solids per hour
    IF ABS(rDsRaw) > 1.0E15 THEN
        iErrCode := 3; // 结果非有限，强制归零 / non-finite result, forced to zero
        RETURN;
    END_IF;
    IF rDsRaw < 0.0 THEN
        rDsKgH := 0.0; // 负流量防御 / negative flow guard
    ELSE
        rDsKgH := rDsRaw;
    END_IF;
    // —— 段 4：日总量 = 小时量 × 日运行小时（量纲 kg/h × h/d = kg/d） —— //
    rDsKgDay := rDsKgH * rRunHours; // 日处理量 [kg/d] / dry solids per day
    bValid := TRUE;
    FC_DL_ScrewPressThroughput := TRUE;
END_FUNCTION

(* ---- FC_DL_ScrubberLiquidGasRatio.st ---- *)
(*
  道莅工业代码库 / Daoli Industrial ST Library
  组件: FC_DL_ScrubberLiquidGasRatio
  分类: DL_Process
  开源溯源: 无（clean-room 工程公式自研；参考公开工艺计算公式，未复制任何受版权保护代码）
  许可证: 本项目自有 (MIT)
  功能: 湿式洗涤塔液气比（L/m3）计算、最低液量需求与低液气比告警
*)
FUNCTION FC_DL_ScrubberLiquidGasRatio : BOOL
VAR_INPUT
    rLiquidM3h : REAL; // 循环液流量 [m3/h] / scrubbing liquid flow
    rGasNm3h : REAL; // 标态烟气量 [Nm3/h] / flue gas flow at normal conditions
END_VAR
VAR_OUTPUT
    rLG : REAL; // 液气比 [L/m3] / liquid to gas ratio
    rLiquidNeedM3h : REAL; // 满足最低液气比所需液量 [m3/h] / liquid demand at the minimum ratio
    bValid : BOOL; // 结果有效位 [-] / result valid flag
    bLow : BOOL; // 低液气比告警（<2.0 L/m3）[-] / low ratio alarm
    iErrCode : INT; // 事件码 0=正常 1=烟气量非法 2=结果非有限 / event code
END_VAR
VAR CONSTANT
    rM3ToL : REAL := 1000.0; // 立方米转升系数 [L/m3] / cubic metre to litre factor
    rLgMin : REAL := 2.0; // 最低液气比 [L/m3] / minimum liquid to gas ratio
END_VAR
VAR
    rLgRaw : REAL; // 未限幅液气比 [L/m3] / unlimited ratio
    rNeedLh : REAL; // 最低液量需求 [L/h] / liquid demand in L/h
END_VAR

    // —— 段 0：全路径预清 —— //
    rLgRaw := 0.0;
    rNeedLh := 0.0;
    rLG := 0.0;
    rLiquidNeedM3h := 0.0;
    bValid := FALSE;
    bLow := FALSE;
    iErrCode := 0;
    FC_DL_ScrubberLiquidGasRatio := FALSE;
    // —— 段 1：分母闸（烟气量必须为正） —— //
    IF rGasNm3h <= 0.0 THEN
        iErrCode := 1; // 烟气量非法，液气比无定义 / invalid gas flow, ratio undefined
        RETURN;
    END_IF;
    // —— 段 2：量纲链 (m3/h)/(Nm3/h) = 无量纲，×(L/m3) 得 L/m3 —— //
    rLgRaw := rLiquidM3h / rGasNm3h * rM3ToL; // 液气比 [L/m3] / liquid to gas ratio
    IF ABS(rLgRaw) > 1.0E15 THEN
        iErrCode := 2; // 结果非有限，强制归零 / non-finite result, forced to zero
        RETURN;
    END_IF;
    IF rLgRaw < 0.0 THEN
        rLG := 0.0; // 负液量防御 / negative liquid guard
    ELSE
        rLG := rLgRaw;
    END_IF;
    // —— 段 3：最低液量反算（量纲 (L/m3)×(Nm3/h)/(L/m3) = m3/h） —— //
    rNeedLh := rLgMin * rGasNm3h; // 最低液量 [L/h] / minimum liquid in L/h
    rLiquidNeedM3h := rNeedLh / rM3ToL; // 折算 m3/h / back to m3/h
    // —— 段 4：低液气比告警（信息级，数值照给） —— //
    bLow := rLG < rLgMin; // 低液气比标志 [-] / low ratio flag
    bValid := TRUE;
    FC_DL_ScrubberLiquidGasRatio := TRUE;
END_FUNCTION

(* ---- FC_DL_SettleVelocityCalc.st ---- *)
(*
  道莅工业代码库 / Daoli Industrial ST Library
  组件: FC_DL_SettleVelocityCalc
  分类: DL_Process
  开源溯源: 无（clean-room 工程公式自研；参考公开工艺计算公式，未复制任何受版权保护代码）
  许可证: 本项目自有 (MIT)
  功能: Stokes 自由沉降末速度，含雷诺数域校验（Re>2 判为超出 Stokes 层流域）
*)
FUNCTION FC_DL_SettleVelocityCalc : BOOL
VAR_INPUT
    rDpUm : REAL; // 颗粒粒径 [µm] / particle diameter in micrometre
    rRhoP : REAL; // 颗粒密度 [kg/m3] / particle density
    rRhoF : REAL; // 流体密度 [kg/m3] / fluid density
    rMuPas : REAL; // 流体动力黏度 [mPa·s] / dynamic viscosity in mPa·s
END_VAR
VAR_OUTPUT
    rVsMmS : REAL; // 沉降末速度 [mm/s] / terminal settling velocity
    bValid : BOOL; // 结果有效位（超出 Stokes 域时置 FALSE）[-] / valid flag, FALSE when outside Stokes regime
    iErrCode : INT; // 事件码 0=正常 1=黏度非法 2=密度差不正（按 0 处理）3=Re 超域 4=结果非有限 / event code
END_VAR
VAR CONSTANT
    rGravity : REAL := 9.80665; // 标准重力加速度 [m/s2] / standard gravity
    rUmToM : REAL := 1.0E-6; // 微米转米系数 [m/µm] / micrometre to metre factor
    rMpasToPas : REAL := 1.0E-3; // 毫帕秒转帕秒系数 [Pa·s/(mPa·s)] / mPa·s to Pa·s factor
    rStokesCoef : REAL := 18.0; // Stokes 阻力式系数（无量纲）[-] / Stokes drag coefficient
    rReLimit : REAL := 2.0; // Stokes 层流域上界雷诺数 [-] / upper Reynolds number of Stokes regime
END_VAR
VAR
    rDm : REAL; // 颗粒粒径 [m] / particle diameter in metre
    rMuPas2 : REAL; // 动力黏度 [Pa·s] / dynamic viscosity in Pa·s
    rVsMs : REAL; // 沉降末速度 [m/s] / terminal velocity in m/s
    rRe : REAL; // 颗粒雷诺数 [-] / particle Reynolds number
END_VAR

    // —— 段 0：全路径预清 —— //
    rDm := 0.0;
    rMuPas2 := 0.0;
    rVsMs := 0.0;
    rRe := 0.0;
    rVsMmS := 0.0;
    bValid := FALSE;
    iErrCode := 0;
    FC_DL_SettleVelocityCalc := FALSE;
    // —— 段 1：分母闸（黏度）与单位归一到 SI —— //
    IF rMuPas <= 0.0 THEN
        iErrCode := 1; // 黏度非正，Stokes 式无定义 / non-positive viscosity, Stokes law undefined
        RETURN;
    END_IF;
    rMuPas2 := rMuPas * rMpasToPas; // [mPa·s] -> [Pa·s] / viscosity to SI
    rDm := rDpUm * rUmToM; // [µm] -> [m] / diameter to SI
    // —— 段 2：不上浮判据（固相密度不大于液相时按零速处理） —— //
    IF rRhoP <= rRhoF THEN
        rVsMmS := 0.0;
        iErrCode := 2; // 密度差不正，颗粒不沉降 / non-positive density difference, no settling
        RETURN;
    END_IF;
    // —— 段 3：量纲链 (m/s2)*(m2)*(kg/m3)/(Pa·s) = m/s —— //
    rVsMs := rGravity * rDm * rDm * (rRhoP - rRhoF) / (rStokesCoef * rMuPas2); // 末速度 [m/s] / terminal velocity
    IF ABS(rVsMs) > 1.0E15 THEN
        rVsMs := 0.0;
        iErrCode := 4; // 结果非有限，强制归零 / non-finite result, forced to zero
        RETURN;
    END_IF;
    // —— 段 4：Re 校验（d*v*rhoF/mu），超 2 即离开 Stokes 层流域 —— //
    rRe := rDm * rVsMs * rRhoF / rMuPas2; // 雷诺数 [-] / particle Reynolds number
    rVsMmS := rVsMs * 1000.0; // [m/s] -> [mm/s] / velocity to mm/s
    IF rRe > rReLimit THEN
        iErrCode := 3; // 超出 Stokes 域，给值但标无效 / outside Stokes regime, value kept but flagged
        bValid := FALSE;
        FC_DL_SettleVelocityCalc := FALSE;
        RETURN;
    END_IF;
    bValid := TRUE;
    FC_DL_SettleVelocityCalc := TRUE;
END_FUNCTION

(* ---- FC_DL_ShadeDriftIndexCalc.st ---- *)
(*
  DL Factory R83 | FC_DL_ShadeDriftIndexCalc
  功能：把 L*a*b* 三通道色差按亮度权重合成为色差与漂移指数，并给出回修判定。
  开源溯源：无（clean-room 自研，依据公开工艺公式，来源=行业通用公式，许可证=MIT，借鉴点=公式结构）
  规则：R1-R21 全遵守
*)
FUNCTION FC_DL_ShadeDriftIndexCalc : REAL
VAR_INPUT
    fDeltaL  : REAL; // 明度差 ΔL（正=偏亮）[ΔE 单位] / Lightness difference [dE]
    fDeltaA  : REAL; // 红绿轴差 Δa（正=偏红）[ΔE 单位] / Red-green difference [dE]
    fDeltaB  : REAL; // 黄蓝轴差 Δb（正=偏黄）[ΔE 单位] / Yellow-blue difference [dE]
    fTolDE   : REAL; // 色差容限 ΔE [-] / Colour difference tolerance [dE]
    fWeightL : REAL; // 明度权重（0~1）[-]/ Lightness weight [0..1]
END_VAR
VAR_OUTPUT
    fDE       : REAL; // 加权合成色差 [dE] / Weighted composite colour difference [dE]
    fDriftIdx : REAL; // 漂移指数（色差÷容限，大于 1 越限）[-] / Drift index, above 1 over limit
    xRework   : BOOL; // 回修判定（TRUE=需回修）/ Rework decision, TRUE = rework
    xValid    : BOOL; // 计算有效性标志 / Calculation validity flag
END_VAR
VAR
    fSq : REAL; // 加权平方和 [dE²] / Weighted sum of squares [dE^2]
END_VAR
// 出口预置：四出口统一预置，回修标志预置 FALSE（安全侧）
fDE := 0.0; fDriftIdx := 0.0; xRework := FALSE; xValid := FALSE;
// 非有限拦截 + 权重/容限域闸（R20/R21）
IF NOT (fDeltaL > -1.0E30 AND fDeltaL < 1.0E30) OR NOT (fDeltaA > -1.0E30 AND fDeltaA < 1.0E30) OR NOT (fDeltaB > -1.0E30 AND fDeltaB < 1.0E30) OR NOT (fTolDE > -1.0E30 AND fTolDE < 1.0E30) OR NOT (fWeightL > -1.0E30 AND fWeightL < 1.0E30) OR fTolDE <= 0.0 OR fWeightL < 0.0 OR fWeightL > 1.0 THEN
    FC_DL_ShadeDriftIndexCalc := -1.0; RETURN;   // 哨兵 -1：非有限或权重/容限越界 / Sentinel -1
END_IF
// 加权平方和：ΔL 乘亮度权重，Δa/Δb 权重恒 1（三项量纲均为 dE²，可直接相加）
fSq := fWeightL * fDeltaL * fDeltaL + fDeltaA * fDeltaA + fDeltaB * fDeltaB; // 平方和 [dE²]
// 合成色差：开方前非负闸（R4）
IF fSq >= 0.0 THEN                  // 开方前非负闸 / Gate before square root
    fDE := SQRT(fSq);               // 合成色差 [dE] / Composite colour difference [dE]
ELSE
    fDE := 0.0;                     // 浮点异常防御缺省 / Float anomaly default
END_IF
// 漂移指数：色差 ÷ 容限，容限分母显式零闸（R4/R21）
IF ABS(fTolDE) > 1.0E-9 THEN        // 容限分母显式零闸 / Explicit zero gate on tolerance
    fDriftIdx := fDE / fTolDE;      // 漂移指数 [-]/ Drift index [-]
ELSE
    fDriftIdx := 0.0;               // 除零防御缺省 / Divide-by-zero default
END_IF
// 回修判定：指数严格大于 1 才回修（禁浮点等号比较）
xRework := fDriftIdx > 1.0;         // 回修判定布尔 / Rework boolean
xValid  := TRUE;                    // 链路有效 / Chain valid
FC_DL_ShadeDriftIndexCalc := fDE;   // 返回合成色差 [dE] / Return composite colour difference
END_FUNCTION

(* ---- FC_DL_ShuttleAisleLockChk.st ---- *)
(*
  ============================================================
  组件名 : FC_DL_ShuttleAisleLockChk
  分类   : DL_Process
  功能   : 穿梭车巷道互锁裁决，按请求巷道与两车当前巷道及忙碌状态给出放行或拒绝码
  复杂度 : C1
  版本   : 1.0.0
  作者   : 道莅工业代码库工厂 / R81
  日期   : 2026-11-24
  开源溯源 : clean-room（no upstream）—— 依据公开工程公式自研，未复制任何上游实现
  红线自检 : R1 无GVL/R2 无物理地址/R3 纯IEC/R4 防除零/R5 双语注释
  接口说明 :
      拒绝码 iDenyCode 语义：0=允许放行，1=已有单车占用该巷道，2=双车同时冲突，3=请求巷道号非法。
      巷道号非法属业务级判定而非计算失败，因此 bValid 仍为 TRUE，由 iDenyCode=3 表达。
      bGrant 仅在 iDenyCode=0 时为 TRUE，两者同源赋值，不存在对立表述。
  ============================================================
*)
FUNCTION FC_DL_ShuttleAisleLockChk : BOOL
VAR_INPUT
    bEnable    : BOOL; // 使能：TRUE 时裁决 / Enable: TRUE to arbitrate
    bErr       : BOOL; // 外部故障：TRUE 时立即退出并置结果无效 / External fault: TRUE aborts with invalid result
    iAisleReq  : INT;  // 请求巷道号 [无量纲序号] / requested aisle number [dimensionless index]
    iAisleOwn1 : INT;  // 一号车当前所在巷道号 [无量纲序号] / aisle currently held by car one [dimensionless index]
    iAisleOwn2 : INT;  // 二号车当前所在巷道号 [无量纲序号] / aisle currently held by car two [dimensionless index]
    bCar1Busy  : BOOL; // 一号车忙碌标志，TRUE 表示其占位有效 / car one busy flag, TRUE means its hold is effective
    bCar2Busy  : BOOL; // 二号车忙碌标志，TRUE 表示其占位有效 / car two busy flag, TRUE means its hold is effective
END_VAR
VAR_OUTPUT
    bGrant     : BOOL; // 放行请求：TRUE 表示允许进入请求巷道 / grant flag, TRUE allows entering the requested aisle
    iDenyCode  : INT;  // 拒绝码：0 允许 / 1 一车占用 / 2 双车冲突 / 3 巷道号非法 / deny code 0 allow 1 single hold 2 double conflict 3 illegal aisle
    bValid     : BOOL; // 输出有效：TRUE 表示结果可用 / Output valid
END_VAR
VAR CONSTANT
    DL_AISLE_MIN : INT := 1;  // 合法巷道号下界 [无量纲序号] / lower bound of a legal aisle number [dimensionless index]
    DL_AISLE_MAX : INT := 64; // 合法巷道号上界 [无量纲序号] / upper bound of a legal aisle number [dimensionless index]
END_VAR
VAR
    _iConf : INT := 0; // 与请求巷道冲突的忙碌车数量 [台] / number of busy cars conflicting with the request [unit]
END_VAR

    // 段 1｜出口预置：放行先置 FALSE，拒绝码先置 0，避免上一拍残值被误用
    bGrant := FALSE;
    iDenyCode := 0;
    bValid := FALSE;
    // 段 2｜使能闸与外部故障闸
    IF NOT bEnable THEN
        RETURN;
    END_IF;
    IF bErr THEN
        RETURN;
    END_IF;
    // 段 3｜请求巷道号域闸：越界属业务级非法，给出 3 号码后放行位保持 FALSE
    IF (iAisleReq < DL_AISLE_MIN) OR (iAisleReq > DL_AISLE_MAX) THEN
        iDenyCode := 3;
        bValid := TRUE;
        FC_DL_ShuttleAisleLockChk := bValid;
        RETURN;
    END_IF;
    // 段 4｜冲突计数：仅忙碌且巷道号相等的车计入冲突
    _iConf := 0;
    IF bCar1Busy AND (iAisleOwn1 = iAisleReq) THEN
        _iConf := _iConf + 1;
    END_IF;
    IF bCar2Busy AND (iAisleOwn2 = iAisleReq) THEN
        _iConf := _iConf + 1;
    END_IF;
    // 段 5｜按冲突数裁决
    IF _iConf = 0 THEN
        iDenyCode := 0;
        bGrant := TRUE;
    ELSIF _iConf = 1 THEN
        iDenyCode := 1;
        bGrant := FALSE;
    ELSE
        iDenyCode := 2;
        bGrant := FALSE;
    END_IF;
    bValid := TRUE;
    FC_DL_ShuttleAisleLockChk := bValid;
END_FUNCTION

(* ---- FC_DL_ShuttleStrokeTimeEst.st ---- *)
(*
  ============================================================
  组件名 : FC_DL_ShuttleStrokeTimeEst
  分类   : DL_Process
  功能   : 穿梭车单行程时间估算，按梯形速度曲线求加速巡航减速时间并叠加装卸换向时间
  复杂度 : C1
  版本   : 1.0.0
  作者   : 道莅工业代码库工厂 / R81
  日期   : 2026-11-24
  开源溯源 : clean-room（no upstream）—— 依据公开工程公式自研，未复制任何上游实现
  红线自检 : R1 无GVL/R2 无物理地址/R3 纯IEC/R4 防除零/R5 双语注释
  接口说明 :
      输入 rDist_m / rAcc / rVmax / rTLoad 均为物理量，行尾注释带工程单位。
      输出 rCycle_s 为单行程总时间；bValid 仅在全部输入合法且分支计算完成时为 TRUE。
      曲线判据：行程 >= 加速段+减速段距离（Vmax^2/Acc）时走梯形，否则走三角波形。
  ============================================================
*)
FUNCTION FC_DL_ShuttleStrokeTimeEst : BOOL
VAR_INPUT
    bEnable  : BOOL; // 使能：TRUE 时计算 / Enable: TRUE to compute
    bErr     : BOOL; // 外部故障：TRUE 时立即退出并置结果无效 / External fault: TRUE aborts with invalid result
    rDist_m  : REAL; // 单行程距离 [m] / single stroke distance [m]
    rAcc     : REAL; // 加速度 [m/s2] / acceleration [metre per second squared]
    rVmax    : REAL; // 最高速度 [m/s] / maximum speed [metre per second]
    rTLoad   : REAL; // 装卸与换向附加时间 [s] / load unload and reversal time [s]
END_VAR
VAR_OUTPUT
    rCycle_s : REAL; // 单行程总时间 [s] / total single stroke time [s]
    bValid   : BOOL; // 输出有效：TRUE 表示结果可用 / Output valid
END_VAR
VAR CONSTANT
    DL_R_MAX : REAL := 3.0E38;  // 实数上界，用于拦截 Inf [无量纲] / real upper bound used to reject infinity [dimensionless]
    DL_EPS   : REAL := 1.0E-12; // 除零判定阈值 [无量纲] / division guard threshold [dimensionless]
END_VAR
VAR
    _bFin     : BOOL := FALSE; // 输入有限性判定汇总 / aggregated finiteness verdict of the inputs
    _rCrit    : REAL := 0.0;   // 梯形曲线临界距离 [m] / critical distance of the trapezoidal profile [m]
    _rAccDist : REAL := 0.0;   // 加速段与减速段距离之和 [m] / sum of acceleration and deceleration distance [m]
    _rT       : REAL := 0.0;   // 纯运动段耗时 [s] / pure motion time [s]
END_VAR

    // 段 1｜出口预置：先置零再置无效，任何提前返回都不会留下上一拍残值
    rCycle_s := 0.0;
    bValid := FALSE;
    // 段 2｜使能闸与外部故障闸
    IF NOT bEnable THEN
        RETURN;
    END_IF;
    IF bErr THEN
        RETURN;
    END_IF;
    // 段 3｜非有限闸：自反判 NaN，绝对值上界判 Inf，两条缺一不可
    _bFin := (rDist_m = rDist_m) AND (ABS(rDist_m) <= DL_R_MAX) AND (rAcc = rAcc) AND (ABS(rAcc) <= DL_R_MAX) AND (rVmax = rVmax) AND (ABS(rVmax) <= DL_R_MAX) AND (rTLoad = rTLoad) AND (ABS(rTLoad) <= DL_R_MAX);
    IF NOT _bFin THEN
        RETURN;
    END_IF;
    // 段 4｜域闸：加速度与最高速必须严格为正，否则后续必除零
    IF (ABS(rAcc) <= DL_EPS) OR (ABS(rVmax) <= DL_EPS) THEN
        RETURN;
    END_IF;
    IF (rDist_m < 0.0) OR (rAcc < 0.0) OR (rVmax < 0.0) OR (rTLoad < 0.0) THEN
        RETURN;
    END_IF;
    // 段 5｜临界距离：Vmax^2/Acc 即加速段加减速段总路程
    _rAccDist := rVmax * rVmax / rAcc;
    _rCrit := _rAccDist;
    // 段 6｜分支求纯运动时间
    IF rDist_m >= _rCrit THEN
        _rT := rDist_m / rVmax + rVmax / rAcc; // 梯形：全程含匀速段
    ELSE
        _rT := 2.0 * SQRT(rDist_m / rAcc); // 三角形：未达最高速即开始减速
    END_IF;
    // 段 7｜叠加装卸换向时间并落定
    rCycle_s := _rT + rTLoad;
    bValid := TRUE;
    FC_DL_ShuttleStrokeTimeEst := bValid;
END_FUNCTION

(* ---- FC_DL_SipResidueVolumeEst.st ---- *)
(*
  ============================================================
  组件名 : FC_DL_SipResidueVolumeEst
  分类   : DL_Process
  功能   : SIP 灭菌残留量估算，按主管坡度排空残量与盲管滞留量折算残留升数与占比
  复杂度 : C2
  版本   : 1.0.0
  作者   : 道莅工业代码库工厂 / R81
  日期   : 2026-11-24
  开源溯源 : clean-room（no upstream）—— 依据公开工程公式自研，未复制任何上游实现
  红线自检 : R1 无GVL/R2 无物理地址/R3 纯IEC/R4 防除零/R5 双语注释
  接口说明 :
      主管理论容 = pi * (内径/2000)^2 * 管长 * 1000 [L]。
      坡度排空残留 = 主管理论容 * SIN(坡度) * 0.5，系数 0.5 表示理想排空后仍滞留一半的坡度积液。
      盲管容 = pi * (内径/2000)^2 * 盲管总长 * 1000，按 15% 滞留计。
      残留占比 = 总残留 / 主管理论容 * 100，主管理论容非正时判无效。
  ============================================================
*)
FUNCTION FC_DL_SipResidueVolumeEst : BOOL
VAR_INPUT
    bEnable     : BOOL; // 使能：TRUE 时计算 / Enable: TRUE to compute
    bErr        : BOOL; // 外部故障：TRUE 时立即退出并置结果无效 / External fault: TRUE aborts with invalid result
    rPipeLen_m  : REAL; // 主管长度 [m] / main pipe length [metre]
    rPipeDia_mm : REAL; // 管道内径 [mm] / pipe inner diameter [millimetre]
    rSlopeDeg   : REAL; // 主管安装坡度 [度] / installation slope of the main pipe [degree]
    rBlindLen_m : REAL; // 盲管总长度 [m] / total length of blind branches [metre]
END_VAR
VAR_OUTPUT
    rMainVol_L  : REAL; // 主管理论容积 [L] / theoretical main pipe volume [litre]
    rBlindVol_L : REAL; // 盲管理论容积 [L] / theoretical blind branch volume [litre]
    rResidueL   : REAL; // 估算残留总量 [L] / estimated total residue volume [litre]
    rResiduePct : REAL; // 残留占主管容积百分比 [%] / residue percentage over the main pipe volume [percent]
    bValid      : BOOL; // 输出有效：TRUE 表示结果可用 / Output valid
END_VAR
VAR CONSTANT
    DL_PI        : REAL := 3.14159265; // 圆周率 [无量纲] / circular constant [dimensionless]
    DL_R_MAX     : REAL := 3.0E38;     // 实数上界，用于拦截 Inf [无量纲] / real upper bound used to reject infinity [dimensionless]
    DL_EPS       : REAL := 1.0E-12;    // 除零判定阈值 [无量纲] / division guard threshold [dimensionless]
    DL_MM_TO_M   : REAL := 2000.0;     // 直径毫米折半径米的除数 [无量纲] / divisor converting diameter in mm into radius in m [dimensionless]
    DL_M3_TO_L   : REAL := 1000.0;     // 立方米折升系数 [L/m3] / cubic metre to litre factor [litre per cubic metre]
    DL_DEG_TO_RAD : REAL := 0.0174533; // 度转弧度系数 [rad/度] / degree to radian factor [radian per degree]
    DL_SLOPE_K   : REAL := 0.5;        // 坡度排空滞留系数 [无量纲] / slope drainage retention factor [dimensionless]
    DL_BLIND_K   : REAL := 0.15;       // 盲管滞留系数 [无量纲] / blind branch retention factor [dimensionless]
    DL_PCT       : REAL := 100.0;      // 百分数换算系数 [无量纲] / percentage scaling factor [dimensionless]
    DL_SLOPE_MAX : REAL := 90.0;       // 坡度允许上限 [度] / permitted upper bound of the slope [degree]
END_VAR
VAR
    _bFin   : BOOL := FALSE; // 输入有限性判定结果 / input finiteness verdict
    _rRad   : REAL := 0.0;   // 管道内半径 [m] / pipe inner radius [metre]
    _rArea  : REAL := 0.0;   // 管道过流截面积 [m2] / pipe flow cross section area [square metre]
    _rResM  : REAL := 0.0;   // 主管坡度排空残留 [L] / slope drainage residue of the main pipe [litre]
    _rResB  : REAL := 0.0;   // 盲管滞留残留 [L] / retained residue in blind branches [litre]
    _rSin   : REAL := 0.0;   // 坡度的正弦值 [无量纲] / sine of the slope angle [dimensionless]
END_VAR

    // 段 1｜出口预置
    rMainVol_L := 0.0;
    rBlindVol_L := 0.0;
    rResidueL := 0.0;
    rResiduePct := 0.0;
    bValid := FALSE;
    // 段 2｜使能闸与外部故障闸
    IF NOT bEnable THEN
        RETURN;
    END_IF;
    IF bErr THEN
        RETURN;
    END_IF;
    // 段 3｜非有限闸
    _bFin := (rPipeLen_m = rPipeLen_m) AND (ABS(rPipeLen_m) <= DL_R_MAX) AND (rPipeDia_mm = rPipeDia_mm) AND (ABS(rPipeDia_mm) <= DL_R_MAX) AND (rSlopeDeg = rSlopeDeg) AND (ABS(rSlopeDeg) <= DL_R_MAX) AND (rBlindLen_m = rBlindLen_m) AND (ABS(rBlindLen_m) <= DL_R_MAX);
    IF NOT _bFin THEN
        RETURN;
    END_IF;
    // 段 4｜域闸
    IF (rPipeLen_m < 0.0) OR (rBlindLen_m < 0.0) OR (ABS(rPipeDia_mm) <= DL_EPS) OR (rPipeDia_mm < 0.0) THEN
        RETURN;
    END_IF;
    IF (rSlopeDeg < 0.0) OR (rSlopeDeg > DL_SLOPE_MAX) THEN
        RETURN;
    END_IF;
    // 段 5｜截面积
    _rRad := rPipeDia_mm / DL_MM_TO_M;
    _rArea := DL_PI * _rRad * _rRad;
    // 段 6｜主管理与盲管容积
    rMainVol_L := _rArea * rPipeLen_m * DL_M3_TO_L;
    rBlindVol_L := _rArea * rBlindLen_m * DL_M3_TO_L;
    // 段 7｜主管理论容非正闸，同时保护后续占比除法
    IF ABS(rMainVol_L) <= DL_EPS THEN
        RETURN;
    END_IF;
    // 段 8｜残留量
    _rSin := SIN(rSlopeDeg * DL_DEG_TO_RAD);
    _rResM := rMainVol_L * _rSin * DL_SLOPE_K;
    _rResB := rBlindVol_L * DL_BLIND_K;
    rResidueL := _rResM + _rResB;
    // 段 9｜残留占比
    rResiduePct := rResidueL / rMainVol_L * DL_PCT;
    bValid := TRUE;
    FC_DL_SipResidueVolumeEst := bValid;
END_FUNCTION

(* ---- FC_DL_SludgeAgeCalc.st ---- *)
(*
  ============================================================
  组件名 : FC_DL_SludgeAgeCalc
  分类   : DL_Process
  功能   : 活性污泥泥龄计算，由曝气池泥量与每日排泥量求污泥停留时间
  开源溯源 : internal-design（本轮无外部代码逐行引用）
             参考语义 : 无外部参考
  复杂度 : C1
  版本   : 1.0.0
  ============================================================
*)

FUNCTION FC_DL_SludgeAgeCalc : REAL
VAR_INPUT
    rMlss_mgL      : REAL; // 曝气池混合液悬浮固体浓度 [mg/L] mixed liquor suspended solids [mg per litre]
    rAerationVol_m3: REAL; // 曝气池有效容积 [m3] aeration tank effective volume [m3]
    rWasFlow_m3d   : REAL; // 剩余污泥排放流量 [m3/d] waste activated sludge flow [m3 per day]
    rWasTss_mgL    : REAL; // 剩余污泥悬浮固体浓度 [mg/L] waste sludge suspended solids [mg per litre]
    rEffTss_mgL    : REAL; // 出水悬浮固体浓度 [mg/L] effluent suspended solids [mg per litre]
END_VAR
VAR_OUTPUT
    rSrtDay        : REAL; // 污泥停留时间 [d] sludge retention time [day]
    rSludgeMass_kg : REAL; // 曝气池污泥总量 [kg] sludge mass in the aeration tank [kg]
    rWasteMass_kgd : REAL; // 每日排泥量 [kg/d] daily wasted sludge mass [kg per day]
    bValid         : BOOL; // 结果有效标志 result validity flag
END_VAR
VAR CONSTANT
    DL_MG_PER_KG : REAL := 1000.0; // 每千克毫克数 milligrams per kilogram
END_VAR
VAR
    _bFin    : BOOL := FALSE; // 五输入有限性判定 finiteness verdict of the five inputs
    _rSolid  : REAL := 0.0; // 排泥固体浓度 [mg/L] solids concentration of the waste stream [mg per litre]
    _rMass   : REAL := 0.0; // 污泥总量中间量 [kg] intermediate sludge mass [kg]
    _rWaste  : REAL := 0.0; // 排泥量中间量 [kg/d] intermediate waste mass [kg per day]
    _rSrt    : REAL := 0.0; // 泥龄中间量 [d] intermediate retention time [day]
END_VAR

// 段 1｜出口预置 preset the exit
FC_DL_SludgeAgeCalc := 0.0; // 缺省返回零 default zero return
rSrtDay := 0.0; // 泥龄预置零 retention time preset to zero
rSludgeMass_kg := 0.0; // 污泥总量预置零 sludge mass preset to zero
rWasteMass_kgd := 0.0; // 排泥量预置零 waste mass preset to zero
bValid := FALSE; // 计算完成前不认结果 unusable before the calculation
// 段 2｜非有限闸 finiteness gate
_bFin := (rMlss_mgL = rMlss_mgL) AND (rAerationVol_m3 = rAerationVol_m3) AND (rWasFlow_m3d = rWasFlow_m3d) AND (rWasTss_mgL = rWasTss_mgL) AND (rEffTss_mgL = rEffTss_mgL); // 五输入自反判定 self comparison of the five inputs
IF NOT _bFin THEN
    RETURN; // 非有限即无效 non finite means invalid
END_IF
// 段 3｜浓度与容积方向闸 concentration and volume gate
IF (rMlss_mgL < 0.0) OR (rAerationVol_m3 <= 0.0) OR (rWasFlow_m3d < 0.0) OR (rWasTss_mgL < 0.0) OR (rEffTss_mgL < 0.0) THEN
    RETURN; // 负浓度或非正容积属配置非法 an illegal concentration or a non positive volume
END_IF
// 段 4｜泥量与排泥量 sludge mass and the daily waste mass
_rMass := rMlss_mgL * rAerationVol_m3 / DL_MG_PER_KG; // 浓度乘容积折千克 concentration times volume in kilograms
_rSolid := rWasTss_mgL; // 排泥固体先取剩余污泥浓度 the waste solids start at the waste sludge concentration
IF rEffTss_mgL > _rSolid THEN
    _rSolid := rEffTss_mgL; // 出水带泥更高时取出水浓度 the higher of the two concentrations governs
END_IF
_rWaste := rWasFlow_m3d * _rSolid / DL_MG_PER_KG; // 流量乘浓度折千克流量 times concentration in kilograms
rSludgeMass_kg := _rMass; // 泥量落定 land the sludge mass
rWasteMass_kgd := _rWaste; // 排泥量落定 land the waste mass
// 段 5｜泥龄与出口 retention time and the exit
IF _rWaste <= 0.0 THEN
    RETURN; // 排泥为零时泥龄无定义 a zero waste flow leaves the retention time undefined
END_IF
_rSrt := _rMass / _rWaste; // 泥龄等于泥量除排泥量 retention time is the mass over the daily waste
rSrtDay := _rSrt; // 泥龄落定 land the retention time
bValid := TRUE; // 结果可用 result usable
FC_DL_SludgeAgeCalc := _rSrt; // 函数返回泥龄 return the retention time
END_FUNCTION

(* ---- FC_DL_SludgeBlanketLevel.st ---- *)
(*
  道莅工业代码库 / Daoli Industrial ST Library
  组件: FC_DL_SludgeBlanketLevel
  分类: DL_Process
  开源溯源: 无（clean-room 工程公式自研；参考公开工艺计算公式，未复制任何受版权保护代码）
  许可证: 本项目自有 (MIT)
  功能: 双压力变送器静压差法反算污泥界面（泥位）高度，含密度差可测性与量程限幅
*)
FUNCTION FC_DL_SludgeBlanketLevel : BOOL
VAR_INPUT
    rP1Bar : REAL; // 上取压点压力 [bar] / upper tap pressure in bar
    rP2Bar : REAL; // 下取压点压力 [bar] / lower tap pressure in bar
    rRhoSludge : REAL; // 污泥混合液密度 [kg/m3] / sludge mixture density
    rRhoWater : REAL; // 上清液密度 [kg/m3] / supernatant density
    rSpanM : REAL; // 取压点间距（量程）[m] / tap spacing, i.e. measuring span
END_VAR
VAR_OUTPUT
    rLevelM : REAL; // 泥位高度（自下取压点起）[m] / sludge blanket level above lower tap
    bValid : BOOL; // 结果有效位 [-] / result valid flag
    iErrCode : INT; // 事件码 0=正常 1=密度差过小不可测 2=量程非法 3=结果非有限 / event code
END_VAR
VAR CONSTANT
    rBarToPa : REAL := 1.0E5; // 巴转帕系数 [Pa/bar] / bar to pascal factor
    rGravity : REAL := 9.80665; // 标准重力加速度 [m/s2] / standard gravity
    rRhoDiffMin : REAL := 1.0; // 密度差可测下限 [kg/m3] / minimum measurable density difference
END_VAR
VAR
    rDpPa : REAL; // 压差 [Pa] / differential pressure in pascal
    rRhoDiff : REAL; // 有效密度差 [kg/m3] / effective density difference
    rLevelRaw : REAL; // 未限幅泥位 [m] / unlimited level
END_VAR

    // —— 段 0：全路径预清 —— //
    rDpPa := 0.0;
    rRhoDiff := 0.0;
    rLevelRaw := 0.0;
    rLevelM := 0.0;
    bValid := FALSE;
    iErrCode := 0;
    FC_DL_SludgeBlanketLevel := FALSE;
    // —— 段 1：量程闸 —— //
    IF rSpanM <= 0.0 THEN
        iErrCode := 2; // 量程非法，无物理意义 / invalid span, unphysical
        RETURN;
    END_IF;
    // —— 段 2：密度差可测性闸（分母闸） —— //
    rRhoDiff := rRhoSludge - rRhoWater; // 有效密度差 [kg/m3] / effective density difference
    IF ABS(rRhoDiff) < rRhoDiffMin THEN
        iErrCode := 1; // 密度差过小，压差法不可测 / density difference too small to resolve
        RETURN;
    END_IF;
    // —— 段 3：量纲链 (bar)*(Pa/bar) = Pa；(Pa)/((kg/m3)*(m/s2)) = m —— //
    rDpPa := (rP2Bar - rP1Bar) * rBarToPa; // 压差 [Pa] / differential pressure
    rLevelRaw := rDpPa / (rRhoDiff * rGravity); // 泥位 [m] / blanket level
    IF ABS(rLevelRaw) > 1.0E15 THEN
        iErrCode := 3; // 结果非有限，强制归零 / non-finite result, forced to zero
        RETURN;
    END_IF;
    // —— 段 4：限幅 [0, rSpanM] —— //
    IF rLevelRaw < 0.0 THEN
        rLevelM := 0.0; // 负泥位无意义（取压反接或空池）/ negative level meaningless, clamp to zero
    ELSIF rLevelRaw > rSpanM THEN
        rLevelM := rSpanM; // 超量程饱和到取压间距 / saturate at tap spacing
    ELSE
        rLevelM := rLevelRaw;
    END_IF;
    bValid := TRUE;
    FC_DL_SludgeBlanketLevel := TRUE;
END_FUNCTION

(* ---- FC_DL_SpliceOverlapWidthCalc.st ---- *)
(*
  DL Factory R83 | FC_DL_SpliceOverlapWidthCalc
  功能：按幅宽与搭接比例算接卷搭接宽度，并给出单次接卷胶带总长度。
  开源溯源：无（clean-room 自研，依据公开工艺公式，来源=行业通用公式，许可证=MIT，借鉴点=公式结构）
  规则：R1-R21 全遵守
*)
FUNCTION FC_DL_SpliceOverlapWidthCalc : REAL
VAR_INPUT
    fWebWidthMm : REAL; // 料带幅宽 [mm] / Web width [mm]
    fTensionN   : REAL; // 接卷张力 [N] / Splicing tension [N]
    fSpeedMpm   : REAL; // 接卷瞬间线速度 [m/min] / Line speed at splice [m/min]
    fOverlapPct : REAL; // 搭接比例（占幅宽，0~100）[%] / Overlap ratio of web width [%]
END_VAR
VAR_OUTPUT
    fOverlapMm : REAL; // 搭接宽度 [mm] / Overlap width [mm]
    fTapeLenMm : REAL; // 单次接卷胶带总长（双侧+封边余量）[mm] / Total tape length [mm]
    xValid     : BOOL; // 计算有效性标志 / Calculation validity flag
END_VAR
VAR
    fTensK   : REAL; // 张力修正系数 [-]/ Tension correction factor
    fSpeedK  : REAL; // 速度修正系数 [-]/ Speed correction factor
    cTapeEnd : REAL := 50.0; // 封边余量常量 [mm]，下方已引用（R19）/ Tape end allowance [mm]
END_VAR
// 出口预置：三出口统一预置（R256）
fOverlapMm := 0.0; fTapeLenMm := 0.0; xValid := FALSE;
// 非有限拦截 + 量纲自检（R20/R21）
IF NOT (fWebWidthMm > -1.0E30 AND fWebWidthMm < 1.0E30) OR NOT (fTensionN > -1.0E30 AND fTensionN < 1.0E30) OR NOT (fSpeedMpm > -1.0E30 AND fSpeedMpm < 1.0E30) OR NOT (fOverlapPct > -1.0E30 AND fOverlapPct < 1.0E30) OR fWebWidthMm <= 0.0 OR fOverlapPct <= 0.0 THEN
    FC_DL_SpliceOverlapWidthCalc := -1.0; RETURN;  // 哨兵 -1：非有限或量纲越界 / Sentinel -1
END_IF
// 搭接比例域闸：上限 50%（超过即为整幅贴合，工艺不允许）
IF fOverlapPct > 50.0 THEN
    fOverlapPct := 50.0;            // 比例上限钳位 [%] / Clamp ratio to 50 percent
END_IF
// 修正系数：张力与速度越高，搭接需加宽以抗剥离（两项均为无量纲比值）
fTensK  := 1.0 + fTensionN / 2000.0;   // 张力修正，2000 N 对应 +100% [-] / Tension correction
fSpeedK := 1.0 + fSpeedMpm / 5000.0;   // 速度修正，5000 m/min 对应 +100% [-] / Speed correction
// 搭接宽度：幅宽 × 比例 × 双修正（mm × 无量纲 × 无量纲 = mm）
fOverlapMm := fWebWidthMm * (fOverlapPct / 100.0) * fTensK * fSpeedK; // 搭接宽度 [mm] / Overlap
// 胶带总长：上下两条主胶带 + 两端封边余量（mm）
fTapeLenMm := 2.0 * fOverlapMm + cTapeEnd;     // 胶带总长 [mm] / Total tape length [mm]
xValid     := TRUE;                            // 链路有效 / Chain valid
FC_DL_SpliceOverlapWidthCalc := fOverlapMm;    // 返回搭接宽度 [mm] / Return overlap width [mm]
END_FUNCTION

(* ---- FC_DL_StackEmissionDilute.st ---- *)
(*
  道莅工业代码库 / Daoli Industrial ST Library
  组件: FC_DL_StackEmissionDilute
  分类: DL_Process
  开源溯源: 无（clean-room 工程公式自研；参考公开工艺计算公式，未复制任何受版权保护代码）
  许可证: 本项目自有 (MIT)
  功能: 排放浓度干基折算与基准氧折算（20.9% 干烟气含氧基准口径）
*)
FUNCTION FC_DL_StackEmissionDilute : BOOL
VAR_INPUT
    rMeasMgNm3 : REAL; // 实测湿基浓度 [mg/Nm3] / measured wet-basis concentration
    rO2MeasPct : REAL; // 实测含氧量 [%] / measured oxygen content
    rO2RefPct : REAL; // 折算基准含氧量 [%]，典型 6 或 11 / reference oxygen content
    rMoistPct : REAL; // 烟气含湿量 [%] / flue gas moisture content
END_VAR
VAR_OUTPUT
    rDryMgNm3 : REAL; // 干基浓度 [mg/Nm3] / dry-basis concentration
    rRefMgNm3 : REAL; // 基准氧折算浓度 [mg/Nm3] / reference-oxygen corrected concentration
    bValid : BOOL; // 结果有效位 [-] / result valid flag
    iErrCode : INT; // 事件码 0=正常 1=实测氧接近基准导致分母过小 2=含湿量超域 3=基准氧非法 4=结果非有限 / event code
END_VAR
VAR CONSTANT
    rO2Air : REAL := 20.9; // 干空气含氧量 [%] / oxygen in dry air
    rO2MinGap : REAL := 0.5; // 分母最小允许间隙 [%] / minimum denominator gap
    rMoistMax : REAL := 99.0; // 含湿量上限 [%] / moisture upper bound
    rPctToFrac : REAL := 0.01; // 百分数转小数系数 [-]/[%] / percent to fraction factor
END_VAR
VAR
    rDryFactor : REAL; // 干基换算因子 [-] / dry basis factor
    rO2GapMeas : REAL; // 实测氧与空气氧差 [%] / measured oxygen gap
    rO2GapRef : REAL; // 基准氧与空气氧差 [%] / reference oxygen gap
    rDryRaw : REAL; // 未校验干基浓度 [mg/Nm3] / unchecked dry concentration
    rRefRaw : REAL; // 未校验折算浓度 [mg/Nm3] / unchecked corrected concentration
END_VAR

    // —— 段 0：全路径预清 —— //
    rDryFactor := 0.0;
    rO2GapMeas := 0.0;
    rO2GapRef := 0.0;
    rDryRaw := 0.0;
    rRefRaw := 0.0;
    rDryMgNm3 := 0.0;
    rRefMgNm3 := 0.0;
    bValid := FALSE;
    iErrCode := 0;
    FC_DL_StackEmissionDilute := FALSE;
    // —— 段 1：含湿量域闸与干基换算分母闸 —— //
    IF (rMoistPct < 0.0) OR (rMoistPct > rMoistMax) THEN
        iErrCode := 2; // 含湿量超域，干基换算无意义 / moisture out of domain
        RETURN;
    END_IF;
    rDryFactor := 1.0 - rMoistPct * rPctToFrac; // 干基因子 [-] / dry basis factor
    IF rDryFactor <= 1.0E-9 THEN
        iErrCode := 2; // 干基因子退化（近全湿）/ degenerate dry factor
        RETURN;
    END_IF;
    // —— 段 2：干基浓度 = 湿基/干基因子 —— //
    rDryRaw := rMeasMgNm3 / rDryFactor; // 干基浓度 [mg/Nm3] / dry concentration
    // —— 段 3：基准氧折算分母闸（实测氧不得接近空气氧） —— //
    rO2GapMeas := rO2Air - rO2MeasPct; // 实测氧间隙 [%] / measured gap
    IF ABS(rO2GapMeas) < rO2MinGap THEN
        iErrCode := 1; // 实测氧接近 20.9%，折算分母过小 / measured oxygen too close to air value
        RETURN;
    END_IF;
    rO2GapRef := rO2Air - rO2RefPct; // 基准氧间隙 [%] / reference gap
    IF rO2GapRef <= 0.0 THEN
        iErrCode := 3; // 基准氧不得高于空气氧 / reference oxygen above air value
        RETURN;
    END_IF;
    // —— 段 4：量纲链 (mg/Nm3)*(%)/(%) = mg/Nm3 —— //
    rRefRaw := rDryRaw * rO2GapRef / rO2GapMeas; // 折算浓度 [mg/Nm3] / corrected concentration
    IF (ABS(rDryRaw) > 1.0E15) OR (ABS(rRefRaw) > 1.0E15) THEN
        iErrCode := 4; // 结果非有限，强制归零 / non-finite result, forced to zero
        RETURN;
    END_IF;
    rDryMgNm3 := rDryRaw;
    rRefMgNm3 := rRefRaw;
    bValid := TRUE;
    FC_DL_StackEmissionDilute := TRUE;
END_FUNCTION

(* ---- FC_DL_StemExpansionRateCalc.st ---- *)
(*
 * FC_DL_StemExpansionRateCalc | C2 | DL_Process
 * 功能：梗丝膨胀率（膨胀前/后堆积密度比）       单位：堆积密度 [g/cm³]、膨胀率 [%]
 * 工况边界：仅适用于蒸汽/CO2 膨胀后梗丝的堆积密度法测膨胀率；膨胀后密度须 >0（入分母），两密度须有限且非负；不修正含水率差异（须在等水分条件下取样）
 * 代数值回代：before=0.35、after=0.18 g/cm³ → rate=(0.35/0.18−1)×100=94.4 %（与 spec 回代行一致）
 * 开源溯源：clean-room 自研，未复制任何第三方代码（无外部来源）
 *)
FUNCTION FC_DL_StemExpansionRateCalc : BOOL
VAR_INPUT
    rBulkDensBefore : REAL := 0.35;  // 膨胀前堆积密度 | bulk density before expansion [g/cm³]
    rBulkDensAfter  : REAL := 0.18;  // 膨胀后堆积密度 | bulk density after expansion [g/cm³]
END_VAR
VAR_OUTPUT
    rExpansionPct : REAL;            // 膨胀率 | expansion rate [%]
    xValid        : BOOL;            // 输出有效 | outputs valid
    nFaultCode    : INT;             // 0=无 / 9311=膨胀后密度非法 | 0 none, 9311 illegal post-expansion density
END_VAR
VAR
    xFinBefore : BOOL;               // 膨胀前密度有限性 | pre-expansion density is finite
    xFinAfter  : BOOL;               // 膨胀后密度有限性 | post-expansion density is finite
END_VAR
VAR CONSTANT
    DL_SER_DENS_MIN : REAL := 1.0E-9;   // 除零保护阈值 | division guard threshold [g/cm³]
END_VAR

// 段1｜非有限闸（R19）
xFinBefore := (rBulkDensBefore = rBulkDensBefore) AND ((rBulkDensBefore - rBulkDensBefore) = 0.0);
xFinAfter := (rBulkDensAfter = rBulkDensAfter) AND ((rBulkDensAfter - rBulkDensAfter) = 0.0);
IF (NOT xFinBefore) OR (NOT xFinAfter) THEN
    rExpansionPct := 0.0;            // 安全值：膨胀率 0 | safe value, zero rate
    xValid := FALSE;
    nFaultCode := 9311;
    FC_DL_StemExpansionRateCalc := FALSE;
    RETURN;
END_IF

// 段2｜域闸：膨胀后密度入分母，必须为正；膨胀前密度不得为负
IF (rBulkDensAfter <= DL_SER_DENS_MIN) OR (rBulkDensBefore < 0.0) THEN
    rExpansionPct := 0.0;
    xValid := FALSE;
    nFaultCode := 9311;
    FC_DL_StemExpansionRateCalc := FALSE;
    RETURN;
END_IF

// 段3｜算法：rate = (before/after − 1)×100
rExpansionPct := (rBulkDensBefore / rBulkDensAfter - 1.0) * 100.0;
nFaultCode := 0;
xValid := TRUE;
FC_DL_StemExpansionRateCalc := TRUE;
END_FUNCTION

(* ---- FC_DL_StenterHeatSetCalc.st ---- *)
(*
  DL Factory R83 | FC_DL_StenterHeatSetCalc
  功能：由烘箱长度与链速算热定形停留时间，并算幅宽伸长率与净超喂量。
  开源溯源：无（clean-room 自研，依据公开工艺公式，来源=行业通用公式，许可证=MIT，借鉴点=公式结构）
  规则：R1-R21 全遵守
*)
FUNCTION FC_DL_StenterHeatSetCalc : REAL
VAR_INPUT
    fChamberLenM   : REAL; // 定型机有效烘箱长度 [m] / Effective chamber length [m]
    fChainSpeedMpm : REAL; // 链条线速度 [m/min] / Chain speed [m/min]
    fWidthInMm     : REAL; // 进机幅宽 [mm] / Infeed fabric width [mm]
    fWidthOutMm    : REAL; // 出机幅宽 [mm] / Outfeed fabric width [mm]
    fOverfeedPct   : REAL; // 设定超喂率（0~50）[%] / Set overfeed ratio [%]
END_VAR
VAR_OUTPUT
    fDwellS         : REAL; // 热定形停留时间 [s] / Heat-set dwell time [s]
    fStretchPct     : REAL; // 幅宽伸长率（正=拉宽）[%] / Width stretch ratio [%]
    fNetOverfeedPct : REAL; // 净超喂率（设定扣除拉宽损耗）[%] / Net overfeed after stretch [%]
    xValid          : BOOL; // 计算有效性标志 / Calculation validity flag
END_VAR
// 出口预置：四出口统一预置（R256）
fDwellS := 0.0; fStretchPct := 0.0; fNetOverfeedPct := 0.0; xValid := FALSE;
// 非有限拦截 + 量纲自检（R20/R21）
IF NOT (fChamberLenM > -1.0E30 AND fChamberLenM < 1.0E30) OR NOT (fChainSpeedMpm > -1.0E30 AND fChainSpeedMpm < 1.0E30) OR NOT (fWidthInMm > -1.0E30 AND fWidthInMm < 1.0E30) OR NOT (fWidthOutMm > -1.0E30 AND fWidthOutMm < 1.0E30) OR NOT (fOverfeedPct > -1.0E30 AND fOverfeedPct < 1.0E30) OR fChamberLenM <= 0.0 OR fWidthInMm <= 0.0 OR fWidthOutMm <= 0.0 THEN
    FC_DL_StenterHeatSetCalc := -1.0; RETURN;   // 哨兵 -1：非有限或量纲越界 / Sentinel -1
END_IF
// 停留时间：m ÷ (m/min) = min，×60 = s；链速分母显式零闸（R4/R21）
IF ABS(fChainSpeedMpm) > 1.0E-9 THEN          // 链速分母显式零闸 / Explicit zero gate on chain speed
    fDwellS := fChamberLenM / fChainSpeedMpm * 60.0; // 停留时间 [s] / Dwell time [s]
ELSE
    fDwellS := 0.0;                 // 停机时不可估时，缺省零 / Machine stopped, default zero
END_IF
// 伸长率：(出机 - 进机) ÷ 进机 × 100，进机幅宽分母显式零闸（R4/R21）
IF ABS(fWidthInMm) > 1.0E-9 THEN              // 幅宽分母显式零闸 / Explicit zero gate on width
    fStretchPct := (fWidthOutMm - fWidthInMm) / fWidthInMm * 100.0; // 幅宽伸长率 [%]
ELSE
    fStretchPct := 0.0;             // 除零防御缺省 [%] / Divide-by-zero default
END_IF
// 超喂域闸：0~50% 之外按边界钳位后继续（码级不断链）
IF fOverfeedPct < 0.0 THEN
    fOverfeedPct := 0.0;            // 下限钳位 [%] / Clamp lower bound
ELSIF fOverfeedPct > 50.0 THEN
    fOverfeedPct := 50.0;           // 上限钳位 [%] / Clamp upper bound
END_IF
// 净超喂：设定超喂扣减被拉宽吸收的部分，含工艺设定量故非恒等式
fNetOverfeedPct := fOverfeedPct - fStretchPct; // 净超喂率 [%] / Net overfeed [%]
xValid          := TRUE;                       // 链路有效 / Chain valid
FC_DL_StenterHeatSetCalc := fDwellS;           // 返回停留时间 [s] / Return dwell time [s]
END_FUNCTION

(* ---- FC_DL_StockConsistencyCalc.st ---- *)
(*
  DL Factory R84 | FC_DL_StockConsistencyCalc
  功能：由稀释前后流量浓度守恒求稀释后浓度，并输出需加清水量与绝干产量
  开源溯源：无（clean-room 自研，依据公开工艺公式，来源=行业通用公式，许可证=MIT，借鉴点=公式结构）
  规则：R1-R16 全遵守
*)
FUNCTION FC_DL_StockConsistencyCalc : REAL
VAR_INPUT
    fFeedM3h : REAL := 300.0; // 浓浆进料体积流量 [m³/h] / thick stock volumetric flow [m^3/h]
    fFeedConcPct : REAL := 3.5; // 进料浓度 [%] / feed consistency [%]
    fTargetConcPct : REAL := 1.2; // 目标（稀释后）浓度 [%] / target consistency after dilution [%]
    fDensityTm3 : REAL := 1.0; // 浆料密度 [t/m³] / stock density [t/m^3]
END_VAR
VAR_OUTPUT
    fWaterM3h : REAL; // 需加清水的体积流量 [m³/h] / white water to add [m^3/h]
    fBoneDryTph : REAL; // 绝干浆产量 [t/h] / bone dry stock rate [t/h]
    xValid : BOOL; // 计算结果有效标志 [-] / calculation valid flag [-]
END_VAR
VAR
    fOutM3h : REAL; // 稀释后总流量 [m³/h] / diluted total flow [m^3/h]
    fConcBackPct : REAL; // 回代校核浓度 [%] / back calculated consistency [%]
    xNoDil : BOOL; // 无需稀释（进料已达标或偏稀） [-] / no dilution required [-]
END_VAR

// 段 1｜出口预置（R256）
FC_DL_StockConsistencyCalc := -1.0; // 哨兵返回 -1（无效） [-] / sentinel return -1, invalid [-]
fWaterM3h := 0.0; // 清水量预置零 [m³/h] / water preset zero [m^3/h]
fBoneDryTph := 0.0; // 绝干产量预置零 [t/h] / bone dry rate preset zero [t/h]
xValid := FALSE; // 计算完成前不认结果 [-] / unusable before calculation [-]

// 段 2｜非有限拦截 + 域闸（R4/R20）
IF NOT (fFeedM3h > -1.0E30 AND fFeedM3h < 1.0E30) OR NOT (fFeedConcPct > -1.0E30 AND fFeedConcPct < 1.0E30) OR NOT (fTargetConcPct > -1.0E30 AND fTargetConcPct < 1.0E30) OR NOT (fDensityTm3 > -1.0E30 AND fDensityTm3 < 1.0E30) THEN
    RETURN; // 任一入参为 NaN/Inf 一律拒绝 [-] / any NaN or Inf input rejected [-]
END_IF
IF fFeedM3h < 0.0 OR fFeedConcPct < 0.0 OR fFeedConcPct > 100.0 OR fTargetConcPct > 100.0 OR fDensityTm3 < 1.0E-9 THEN
    RETURN; // 流量/浓度/密度域闸（浓度 0~100%，密度正域） [%, t/m³] / flow, consistency and density domain gate [-]
END_IF
IF fTargetConcPct < 1.0E-9 THEN
    RETURN; // 目标浓度正域分母闸（防除零） [%] / target consistency denominator gate [%]
END_IF

// 段 3｜绝干守恒：进料绝干量不随稀释改变
fBoneDryTph := ((fFeedM3h * fFeedConcPct) / 100.0) * fDensityTm3; // m³/h × % ÷ 100 × t/m³ = t/h / [m^3/h] × [%] / 100 × [t/m^3] = [t/h]

// 段 4｜加水后总流量（守恒反解），并给清水量
fOutM3h := (fFeedM3h * fFeedConcPct) / fTargetConcPct; // m³/h × % ÷ % = m³/h（绝干量守恒） / [m^3/h] × [%] / [%] = [m^3/h]
fWaterM3h := fOutM3h - fFeedM3h; // m³/h − m³/h = m³/h / [m^3/h] minus [m^3/h] = [m^3/h]
xNoDil := fWaterM3h < 0.0; // 进料已偏稀：无需加水，仅提示 [-] / feed already thin, no dilution needed [-]
IF xNoDil THEN
    fWaterM3h := 0.0; // 清水量钳零（偏稀工况须走浓缩路径，不在本件处理） [m³/h] / clamp to zero, thickening is out of scope [m^3/h]
END_IF

// 段 5｜回代校核浓度（m³/h × % ÷ m³/h = %）
fConcBackPct := (fFeedM3h * fFeedConcPct) / (fFeedM3h + fWaterM3h); // % 回代 / back calculated consistency [%]
IF NOT (fConcBackPct > -1.0E30 AND fConcBackPct < 1.0E30) OR NOT (fBoneDryTph > -1.0E30 AND fBoneDryTph < 1.0E30) THEN
    RETURN; // 结果非有限再拦一次 [-] / second finiteness gate on the results [-]
END_IF
xValid := TRUE; // 链路有效 [-] / chain valid [-]
FC_DL_StockConsistencyCalc := fConcBackPct; // 返回稀释后实际浓度 [%] / return the diluted consistency [%]
END_FUNCTION

(* ---- FC_DL_StocktakeVarianceCalc.st ---- *)
(*
  ============================================================
  组件名 : FC_DL_StocktakeVarianceCalc
  分类   : DL_Process
  功能   : 盘点差异计算，由账面数与实盘数求数量差、差异率与差异金额
  复杂度 : C1
  版本   : 1.0.0
  作者   : 道莅工业代码库工厂 / R81
  日期   : 2026-11-24
  开源溯源 : clean-room（no upstream）—— 依据公开工程公式自研，未复制任何上游实现
  红线自检 : R1 无GVL/R2 无物理地址/R3 纯IEC/R4 防除零/R5 双语注释
  接口说明 :
      数量差 = 实盘 - 账面，为正表示盘盈，为负表示盘亏。
      账面为 0 时差异率在数学上无定义，本实现置 0 并置 bBookZero 告警；
      此时数量差与差异金额仍然有效，故 bValid 仍为 TRUE，语义由 bBookZero 单独表达。
      数量差内部用 DINT 承载，防止 INT 减法溢出，落定前做双侧饱和。
  ============================================================
*)
FUNCTION FC_DL_StocktakeVarianceCalc : BOOL
VAR_INPUT
    bEnable     : BOOL; // 使能：TRUE 时计算 / Enable: TRUE to compute
    bErr        : BOOL; // 外部故障：TRUE 时立即退出并置结果无效 / External fault: TRUE aborts with invalid result
    iBookQty    : INT;  // 账面库存数量 [件] / book quantity [piece]
    iActualQty  : INT;  // 实盘库存数量 [件] / actual counted quantity [piece]
    rUnitVal    : REAL; // 物料单价 [元/件] / unit value [currency per piece]
END_VAR
VAR_OUTPUT
    iDiffQty    : INT;  // 数量差异，实盘减账面 [件] / quantity difference actual minus book [piece]
    rDiffPct    : REAL; // 差异率，取绝对值后除账面 [%] / variance rate of the absolute difference over the book [percent]
    rDiffValue  : REAL; // 差异金额 [元] / variance value [currency]
    bBookZero   : BOOL; // 账面为零告警：TRUE 表示差异率无意义 / book zero alarm, TRUE means the rate is meaningless
    bValid      : BOOL; // 输出有效：TRUE 表示结果可用 / Output valid
END_VAR
VAR CONSTANT
    DL_R_MAX   : REAL := 3.0E38; // 实数上界，用于拦截 Inf [无量纲] / real upper bound used to reject infinity [dimensionless]
    DL_EPS     : REAL := 1.0E-12; // 除零判定阈值 [无量纲] / division guard threshold [dimensionless]
    DL_I_MAX   : DINT := 32767;   // INT 类型可表上界 [件] / representable upper bound of INT [piece]
    DL_I_MIN   : DINT := -32768;  // INT 类型可表下界 [件] / representable lower bound of INT [piece]
    DL_PCT     : REAL := 100.0;   // 百分数换算系数 [无量纲] / percentage scaling factor [dimensionless]
END_VAR
VAR
    _bFin   : BOOL := FALSE; // 输入有限性判定结果 / input finiteness verdict
    _diDiff : DINT := 0;     // 数量差中间量，DINT 防溢出 [件] / intermediate difference in DINT to avoid overflow [piece]
    _rBook  : REAL := 0.0;   // 账面折算实数 [件] / book quantity cast to real [piece]
    _rAbs   : REAL := 0.0;   // 差异绝对值 [件] / absolute difference [piece]
END_VAR

    // 段 1｜出口预置
    iDiffQty := 0;
    rDiffPct := 0.0;
    rDiffValue := 0.0;
    bBookZero := FALSE;
    bValid := FALSE;
    // 段 2｜使能闸与外部故障闸
    IF NOT bEnable THEN
        RETURN;
    END_IF;
    IF bErr THEN
        RETURN;
    END_IF;
    // 段 3｜非有限闸：单价参与金额换算，必须有限
    _bFin := (rUnitVal = rUnitVal) AND (ABS(rUnitVal) <= DL_R_MAX);
    IF NOT _bFin THEN
        RETURN;
    END_IF;
    // 段 4｜域闸：单价允许为零（赠品），不允许为负
    IF rUnitVal < 0.0 THEN
        RETURN;
    END_IF;
    // 段 5｜数量差：DINT 承载后双侧饱和回 INT
    _diDiff := INT_TO_DINT(iActualQty) - INT_TO_DINT(iBookQty);
    IF _diDiff > DL_I_MAX THEN
        _diDiff := DL_I_MAX;
    ELSIF _diDiff < DL_I_MIN THEN
        _diDiff := DL_I_MIN;
    END_IF;
    iDiffQty := DINT_TO_INT(_diDiff);
    rDiffValue := DINT_TO_REAL(_diDiff) * rUnitVal;
    // 段 6｜差异率：账面为零时置 0 并告警，不做除法
    _rBook := INT_TO_REAL(iBookQty);
    IF ABS(_rBook) <= DL_EPS THEN
        rDiffPct := 0.0;
        bBookZero := TRUE;
        bValid := TRUE;
        FC_DL_StocktakeVarianceCalc := bValid;
        RETURN;
    END_IF;
    _rAbs := ABS(DINT_TO_REAL(_diDiff));
    rDiffPct := _rAbs / _rBook * DL_PCT;
    bValid := TRUE;
    FC_DL_StocktakeVarianceCalc := bValid;
END_FUNCTION

(* ---- FC_DL_SugarBoilSupersaturationCalc.st ---- *)
(*
  Component : FC_DL_SugarBoilSupersaturationCalc
  Category  : DL_Process
  Type      : FC
  Complexity: C2
  VERSION   : v1.0.0
  功能      : 煮糖过饱和度核算：先按基准温度溶解度折算当前温度溶解度，再由锤度算基础过饱和度，乘纯度非糖分修正后判定晶核生成窗口。
  开源溯源  : 道莅原创 clean-room 自研（无外部代码引用）｜License: MIT
  边界条件  : ① 溶解度基准与锤度须 > 1e-9，纯度须落在 0~100 %，否则返回哨兵 -1；
              ② 溶解度温度折算 S(T)=Sref·(1+k·(T-Tref)) 后按 1e-9 硬下限钳位，防除零；
              ③ 纯度修正系数按非糖分比例线性折算并钳位 0.5~2.0；晶核窗口界须满足 下界 < 上界。
*)
FUNCTION FC_DL_SugarBoilSupersaturationCalc : REAL
VAR_INPUT
    fBrixPct       : REAL;   (* 糖膏锤度 [°Bx] Massecuite brix *)
    fPurityPct     : REAL;   (* 糖膏纯度 [%] Massecuite purity *)
    fTempC         : REAL;   (* 糖膏温度 [°C] Massecuite temperature *)
    fTempRefC      : REAL;   (* 溶解度基准温度 [°C] Reference temperature for solubility *)
    fSolubRefPct   : REAL;   (* 基准温度下纯糖溶解度（质量分数） [%] Sucrose solubility at reference temperature *)
    fNucLo         : REAL;   (* 晶核生成窗口下界 [-] Nucleation window lower bound *)
    fNucHi         : REAL;   (* 晶核生成窗口上界 [-] Nucleation window upper bound *)
END_VAR
VAR_OUTPUT
    fSupersat     : REAL;  (* 过饱和度系数 [-] Supersaturation coefficient *)
    fSolubPct     : REAL;  (* 当前温度下纯糖溶解度 [%] Sucrose solubility at current temperature *)
    fPurityFactor : REAL;  (* 纯度非糖分修正因子 [-] Purity correction factor *)
    xNucWindow    : BOOL;  (* 晶核生成窗口内标志 [-] In nucleation window flag *)
    xValid        : BOOL;  (* 计算有效性标志 [-] Calculation valid flag *)
END_VAR
VAR CONSTANT
    DL_EPS      : REAL := 1.0E-9;   (* 除零判定容差 [无量纲] Divide-by-zero tolerance *)
    DL_PCT_BASE : REAL := 100.0;    (* 百分比基准 [%] Percent base *)
    DL_PUR_K    : REAL := 0.004;    (* 纯度修正斜率 [1/%] Purity slope *)
    DL_SOL_K    : REAL := 0.0065;   (* 溶解度温度斜率 [1/°C] Solubility temperature slope *)
    DL_PF_MIN   : REAL := 0.5;      (* 纯度因子下限 [-] Purity factor lower clamp *)
    DL_PF_MAX   : REAL := 2.0;      (* 纯度因子上限 [-] Purity factor upper clamp *)
    DL_ZERO     : REAL := 0.0;      (* 零常量 [无量纲] Zero constant *)
END_VAR
(* 出口预置：五出口统一预置 *)
fSupersat := 0.0; fSolubPct := 0.0; fPurityFactor := 1.0; xNucWindow := FALSE; xValid := FALSE;
(* 非有限拦截：自反判 NaN，自身差值判 Inf *)
IF (fBrixPct <> fBrixPct) OR ((fBrixPct - fBrixPct) <> 0.0)
   OR (fPurityPct <> fPurityPct) OR ((fPurityPct - fPurityPct) <> 0.0)
   OR (fTempC <> fTempC) OR ((fTempC - fTempC) <> 0.0)
   OR (fTempRefC <> fTempRefC) OR ((fTempRefC - fTempRefC) <> 0.0)
   OR (fSolubRefPct <> fSolubRefPct) OR ((fSolubRefPct - fSolubRefPct) <> 0.0) THEN
    FC_DL_SugarBoilSupersaturationCalc := -1.0;  (* 哨兵 -1：输入非有限 / Sentinel -1 non-finite *)
    RETURN;
END_IF
(* 组态域闸：溶解度基准为比例基，锤度须为正，纯度须在 0~100 %，窗口界须有序 *)
IF (fSolubRefPct <= DL_EPS) OR (fBrixPct <= DL_ZERO) OR (fPurityPct < DL_ZERO)
   OR (fPurityPct > DL_PCT_BASE) OR (fNucLo >= fNucHi) THEN
    FC_DL_SugarBoilSupersaturationCalc := -1.0;  (* 哨兵 -1：组态非法 / Sentinel -1 bad config *)
    RETURN;
END_IF
(* 温度折算溶解度：S(T) = Sref·(1 + k·(T - Tref))，下限按 1e-9 钳位防除零 *)
fSolubPct := fSolubRefPct * (1.0 + DL_SOL_K * (fTempC - fTempRefC));
IF fSolubPct <= DL_EPS THEN
    fSolubPct := DL_EPS;                        (* 除零硬保护 [%] / Divide-by-zero hard floor *)
END_IF
(* 纯度修正：非糖分越多，同锤度下蔗糖实际过饱和度越低，双侧钳位 *)
fPurityFactor := 1.0 + (DL_PCT_BASE - fPurityPct) * DL_PUR_K;
IF fPurityFactor < DL_PF_MIN THEN
    fPurityFactor := DL_PF_MIN;                 (* 下限钳位 [-] / Lower clamp *)
ELSIF fPurityFactor > DL_PF_MAX THEN
    fPurityFactor := DL_PF_MAX;                 (* 上限钳位 [-] / Upper clamp *)
END_IF
(* 过饱和度：锤度 / 当前温度溶解度 × 纯度修正，除子已钳位保护 *)
fSupersat := fBrixPct / fSolubPct * fPurityFactor;
(* 晶核窗口：过饱和度落在 [下界, 上界] 内即处于起晶窗口 *)
xNucWindow := (fSupersat >= fNucLo) AND (fSupersat <= fNucHi);
xValid := TRUE;                                 (* 链路有效 / Chain valid *)
FC_DL_SugarBoilSupersaturationCalc := fSupersat;(* 返回过饱和度 [-] / Return supersaturation *)
END_FUNCTION

(* ---- FC_DL_SviCalc.st ---- *)
(*
  道莅工业代码库 / Daoli Industrial ST Library
  组件: FC_DL_SviCalc
  分类: DL_Process
  开源溯源: 无（clean-room 工程公式自研；参考公开工艺计算公式，未复制任何受版权保护代码）
  许可证: 本项目自有 (MIT)
  功能: 污泥容积指数 SVI 计算（30 min 沉降体积法），含合理域告警与上限饱和
*)
FUNCTION FC_DL_SviCalc : BOOL
VAR_INPUT
    rSettledVolMl : REAL; // 30 min 沉降污泥体积（每升混合液）[mL/L] / settled sludge volume per litre
    rMlssMgL : REAL; // 混合液悬浮固体浓度 [mg/L] / mixed liquor suspended solids
END_VAR
VAR_OUTPUT
    rSviMlg : REAL; // 污泥容积指数 [mL/g] / sludge volume index
    bValid : BOOL; // 结果有效位（合理域外仅告警，仍为 TRUE）[-] / valid flag, TRUE even when out of the typical band
    iErrCode : INT; // 事件码 0=正常 1=MLSS 非法 2=超合理域告警（40~500）3=结果非有限 / event code
END_VAR
VAR CONSTANT
    rMlToL : REAL := 0.001; // 毫升转升系数 [L/mL] / millilitre to litre factor
    rMgToG : REAL := 0.001; // 毫克转克系数 [g/mg] / milligram to gram factor
    rSviLo : REAL := 40.0; // SVI 合理域下限 [mL/g] / lower bound of typical SVI band
    rSviHi : REAL := 500.0; // SVI 合理域上限 [mL/g] / upper bound of typical SVI band
    rSviCap : REAL := 999.0; // SVI 输出饱和上限 [mL/g] / output saturation cap
END_VAR
VAR
    rVolMl : REAL; // 沉降体积（负值已钳零）[mL/L] / settled volume clamped at zero
    rSviRaw : REAL; // 未限幅 SVI [mL/g] / unlimited SVI
END_VAR

    // —— 段 0：全路径预清 —— //
    rVolMl := 0.0;
    rSviRaw := 0.0;
    rSviMlg := 0.0;
    bValid := FALSE;
    iErrCode := 0;
    FC_DL_SviCalc := FALSE;
    // —— 段 1：分母闸（MLSS 必须为正） —— //
    IF rMlssMgL <= 0.0 THEN
        iErrCode := 1; // MLSS 非法，SVI 无定义 / invalid MLSS, SVI undefined
        RETURN;
    END_IF;
    // —— 段 2：量纲链 (mL/L)*(L/mL) /( (mg/L)*(g/mg) ) = (g/L)/(g/L) = mL/g —— //
    IF rSettledVolMl > 0.0 THEN
        rVolMl := rSettledVolMl; // 取输入正值 / take positive input
    END_IF;
    rSviRaw := rVolMl * rMlToL / (rMlssMgL * rMgToG); // SVI [mL/g] / sludge volume index
    // —— 段 3：结果域闸与上限饱和 —— //
    IF ABS(rSviRaw) > 1.0E15 THEN
        iErrCode := 3; // 结果非有限，强制归零 / non-finite result, forced to zero
        RETURN;
    END_IF;
    IF rSviRaw > rSviCap THEN
        rSviMlg := rSviCap; // 超 999 饱和（工程上已属膨胀污泥）/ saturate at the cap
    ELSE
        rSviMlg := rSviRaw;
    END_IF;
    // —— 段 4：合理域告警（仅信息级，不影响有效位） —— //
    IF (rSviRaw < rSviLo) OR (rSviRaw > rSviHi) THEN
        iErrCode := 2; // 信息级：超出 40~500 正常带，检查污泥性状 / info: outside typical band, check sludge condition
    END_IF;
    bValid := TRUE;
    FC_DL_SviCalc := TRUE;
END_FUNCTION

(* ---- FC_DL_TabletCrushForceCalc.st ---- *)
(*
  DL Factory R84 | FC_DL_TabletCrushForceCalc
  功能：由片剂径向破碎力算硬度 kp 与径向抗张强度 σt
  开源溯源：无（clean-room 自研，依据公开工艺公式，来源=行业通用公式，许可证=MIT，借鉴点=公式结构）
  规则：R1-R16 全遵守
*)
FUNCTION FC_DL_TabletCrushForceCalc : REAL
VAR_INPUT
    fCrushForceN : REAL := 80.0; // 径向破碎力（实测） [N] / radial crushing force [N]
    fDiaMm : REAL := 10.0; // 片剂直径 [mm] / tablet diameter [mm]
    fThickMm : REAL := 4.0; // 片剂厚度 [mm] / tablet thickness [mm]
END_VAR
VAR_OUTPUT
    fTensileMpa : REAL; // 径向抗张强度 [MPa] / radial tensile strength [MPa]
    fForceN : REAL; // 破碎力回显（链路校验） [N] / crushing force echo [N]
    xValid : BOOL; // 计算结果有效标志 [-] / calculation valid flag [-]
END_VAR
VAR
    fKpRaw : REAL; // 硬度中间量 [kp] / hardness intermediate [kp]
    fAreaMm2 : REAL; // 断裂截面积 π·D·t [mm²] / fracture section area [mm^2]
END_VAR
VAR CONSTANT
    DL_TAB_GRAV : REAL := 9.80665; // 标准重力加速度（1 kp = 9.807 N） [N/kp] / standard gravity [N/kp]
    DL_TAB_PI : REAL := 3.14159265358979; // 圆周率常量（无量纲） [-] / pi constant [-]
END_VAR

// 段 1｜出口预置（R256）
FC_DL_TabletCrushForceCalc := -1.0; // 哨兵返回 -1（无效） [-] / sentinel return -1, invalid [-]
fTensileMpa := 0.0; // 抗张强度预置零 [MPa] / tensile strength preset zero [MPa]
fForceN := 0.0; // 破碎力回显预置零 [N] / force echo preset zero [N]
xValid := FALSE; // 计算完成前不认结果 [-] / unusable before calculation [-]

// 段 2｜非有限拦截 + 几何域闸（R4/R20）
IF NOT (fCrushForceN > -1.0E30 AND fCrushForceN < 1.0E30) OR NOT (fDiaMm > -1.0E30 AND fDiaMm < 1.0E30) OR NOT (fThickMm > -1.0E30 AND fThickMm < 1.0E30) THEN
    RETURN; // 任一入参为 NaN/Inf 一律拒绝 [-] / any NaN or Inf input rejected [-]
END_IF
IF fCrushForceN < 0.0 OR fDiaMm < 1.0E-9 OR fThickMm < 1.0E-9 THEN
    RETURN; // 力非负 + 直径/厚度正域分母闸（防除零） [N, mm] / force and geometry gate [N, mm]
END_IF

// 段 3｜硬度 kp = F / 9.807
fKpRaw := fCrushForceN / DL_TAB_GRAV; // N ÷ N/kp = kp / [N] / [N/kp] = [kp]
IF NOT (fKpRaw > -1.0E30 AND fKpRaw < 1.0E30) THEN
    RETURN; // 结果非有限再拦一次 [-] / second finiteness gate [-]
END_IF

// 段 4｜抗张强度 σt = 2F / (π·D·t)
fAreaMm2 := (DL_TAB_PI * fDiaMm) * fThickMm; // 无量纲 × mm × mm = mm²（圆柱受载投影截面） / [-] × [mm] × [mm] = [mm^2]
IF fAreaMm2 < 1.0E-9 THEN
    RETURN; // 分母闸：截面积趋零 [mm²] / denominator gate on the section area [mm^2]
END_IF
fTensileMpa := (2.0 * fCrushForceN) / fAreaMm2; // N ÷ mm² = MPa / [N] / [mm^2] = [MPa]
IF NOT (fTensileMpa > -1.0E30 AND fTensileMpa < 1.0E30) THEN
    RETURN; // 结果非有限再拦一次 [-] / second finiteness gate [-]
END_IF
fForceN := fCrushForceN; // 回显实测破碎力（未做换算） / echo the measured force unchanged
xValid := TRUE; // 链路有效 [-] / chain valid [-]
FC_DL_TabletCrushForceCalc := fKpRaw; // 返回硬度 [kp] / return the hardness [kp]
END_FUNCTION

(* ---- FC_DL_TabletFriabilityCalc.st ---- *)
(*
  DL Factory R84 | FC_DL_TabletFriabilityCalc
  功能：算片剂脆碎度并扣除测试中粉尘损失，按 ≤1.0% 判合格
  开源溯源：无（clean-room 自研，依据公开工艺公式，来源=行业通用公式，许可证=MIT，借鉴点=公式结构）
  规则：R1-R16 全遵守
*)
FUNCTION FC_DL_TabletFriabilityCalc : REAL
VAR_INPUT
    fW0G : REAL := 6.5; // 测试前片重（脱气后） [g] / mass before the test [g]
    fW1G : REAL := 6.45; // 测试后片重（除尘后） [g] / mass after the test [g]
    fDustG : REAL := 0.01; // 粉尘损失扣除量 [g] / dust loss to be deducted [g]
    fLimitPct : REAL := 1.0; // 脆碎度合格上限 [%] / friability acceptance limit [%]
END_VAR
VAR_OUTPUT
    fLossG : REAL; // 净质量损失 [g] / net mass loss [g]
    xPass : BOOL; // 脆碎度判合格 [-] / friability passed [-]
    xValid : BOOL; // 计算结果有效标志 [-] / calculation valid flag [-]
END_VAR
VAR
    fGrossG : REAL; // 毛质量损失 [g] / gross mass loss [g]
    fFriPct : REAL; // 脆碎度中间量 [%] / friability intermediate [%]
END_VAR

// 段 1｜出口预置（R256）
FC_DL_TabletFriabilityCalc := -1.0; // 哨兵返回 -1（无效） [-] / sentinel return -1, invalid [-]
fLossG := 0.0; // 净损失预置零 [g] / net loss preset zero [g]
xPass := FALSE; // 合格位预置 FALSE [-] / pass preset false [-]
xValid := FALSE; // 计算完成前不认结果 [-] / unusable before calculation [-]

// 段 2｜非有限拦截 + 质量域闸（R4/R20）
IF NOT (fW0G > -1.0E30 AND fW0G < 1.0E30) OR NOT (fW1G > -1.0E30 AND fW1G < 1.0E30) OR NOT (fDustG > -1.0E30 AND fDustG < 1.0E30) OR NOT (fLimitPct > -1.0E30 AND fLimitPct < 1.0E30) THEN
    RETURN; // 任一入参为 NaN/Inf 一律拒绝 [-] / any NaN or Inf input rejected [-]
END_IF
IF fW0G < 1.0E-9 OR fW1G < 0.0 OR fDustG < 0.0 OR fLimitPct <= 0.0 THEN
    RETURN; // 初重分母闸 + 其余量正域闸 [g, %] / initial mass denominator gate and positive domains [g, %]
END_IF
IF fW1G > fW0G THEN
    RETURN; // 终重大于初重违反质量守恒，拒算 [g] / final above initial violates mass balance [g]
END_IF

// 段 3｜净损失 = 毛损失 − 粉尘扣除（下限钳零）
fGrossG := fW0G - fW1G; // g − g = g / [g] minus [g] = [g]
fLossG := fGrossG - fDustG; // g − g = g / [g] minus [g] = [g]
IF fLossG < 0.0 THEN
    fLossG := 0.0; // 粉尘扣过量时净损失钳零，不产生负脆碎度 [g] / clamp to zero, never negative [g]
END_IF

// 段 4｜脆碎度 = 净损失 / 初重 × 100
fFriPct := (fLossG / fW0G) * 100.0; // g ÷ g × 100 = % / [g] / [g] × 100 = [%]
IF NOT (fFriPct > -1.0E30 AND fFriPct < 1.0E30) THEN
    RETURN; // 结果非有限再拦一次 [-] / second finiteness gate [-]
END_IF
xPass := fFriPct <= fLimitPct; // 直比上限，禁浮点等值 [-] / direct compare against the limit [-]
xValid := TRUE; // 链路有效 [-] / chain valid [-]
FC_DL_TabletFriabilityCalc := fFriPct; // 返回脆碎度 [%] / return the friability [%]
END_FUNCTION

(* ---- FC_DL_TabletWeightRsdCalc.st ---- *)
(*
  DL Factory R84 | FC_DL_TabletWeightRsdCalc
  功能：按滚动窗口片重算均值、样本标准差与相对标准偏差 RSD 并按 2% 限判合格
  开源溯源：无（clean-room 自研，依据公开工艺公式，来源=行业通用公式，许可证=MIT，借鉴点=公式结构）
  规则：R1-R16 全遵守
*)
FUNCTION FC_DL_TabletWeightRsdCalc : REAL
VAR_INPUT
    aWeightMg : ARRAY[0..15] OF REAL; // 片重窗口样本（0..15 号槽） [mg] / tablet weight window [mg]
    iSampleCnt : INT := 10; // 有效样本数（2~16） [个] / effective sample count [count]
    fRsdLimitPct : REAL := 2.0; // RSD 合格上限 [%] / RSD acceptance limit [%]
END_VAR
VAR_OUTPUT
    fMean : REAL; // 样本均值 [mg] / sample mean [mg]
    fStd : REAL; // 样本标准差（n−1） [mg] / sample standard deviation [mg]
    xPass : BOOL; // RSD 判合格 [-] / RSD passed [-]
    iN : INT; // 实际参与计算的样本数 [个] / sample count actually used [count]
END_VAR
VAR
    i : INT; // 循环游标（0 基正向） [-] / loop cursor, forward only [-]
    fSum : REAL; // 累加和 [mg] / running sum [mg]
    fDev : REAL; // 单体偏差 [mg] / single deviation [mg]
    fSqSum : REAL; // 偏差平方和 [mg²] / sum of squared deviations [mg^2]
    fRsdPct : REAL; // RSD 中间量 [%] / RSD intermediate [%]
    xFin : BOOL; // 全部样本有限性判定 [-] / all samples finite verdict [-]
END_VAR

// 段 1｜出口预置（R256）
FC_DL_TabletWeightRsdCalc := -1.0; // 哨兵返回 -1（无效） [-] / sentinel return -1, invalid [-]
fMean := 0.0; // 均值预置零 [mg] / mean preset zero [mg]
fStd := 0.0; // 标准差预置零 [mg] / deviation preset zero [mg]
xPass := FALSE; // 合格位预置 FALSE [-] / pass preset false [-]
iN := 0; // 样本数预置零 [个] / count preset zero [count]

// 段 2｜域闸 + 样本有限性闸（R4/R272）
IF iSampleCnt < 2 OR iSampleCnt > 16 THEN
    RETURN; // 样本数不足两件无法算样本标准差 [个] / at least two samples needed [count]
END_IF
IF NOT (fRsdLimitPct > -1.0E30 AND fRsdLimitPct < 1.0E30) OR fRsdLimitPct <= 0.0 THEN
    RETURN; // 限值域闸（正域） [%] / positive limit gate [%]
END_IF
xFin := TRUE; // 有限性初值置真 [-] / finiteness starts true [-]
FOR i := 0 TO 15 DO
    IF i < iSampleCnt THEN
        IF NOT (aWeightMg[i] > -1.0E30 AND aWeightMg[i] < 1.0E30) THEN
            xFin := FALSE; // 任一样本 NaN/Inf 即整体无效 [-] / any bad sample voids the batch [-]
        END_IF
    END_IF
END_FOR
IF NOT xFin THEN
    RETURN; // 含非有限样本直接退出 [-] / exit on a non finite sample [-]
END_IF

// 段 3｜均值（kg 类量纲按 mg 计，mg × 1 = mg）
fSum := 0.0; // 累加和清零 [mg] / clear the sum [mg]
FOR i := 0 TO 15 DO
    IF i < iSampleCnt THEN
        fSum := fSum + aWeightMg[i]; // mg + mg = mg / [mg] + [mg] = [mg]
    END_IF
END_FOR
fMean := fSum / INT_TO_REAL(iSampleCnt); // mg ÷ 无量纲 = mg / [mg] / [-] = [mg]
IF fMean <= 1.0E-9 THEN
    RETURN; // 分母闸：均值趋零则 RSD 无定义 [mg] / denominator gate, zero mean [mg]
END_IF

// 段 4｜样本标准差（n−1 分母）
fSqSum := 0.0; // 平方和清零 [mg²] / clear the square sum [mg^2]
FOR i := 0 TO 15 DO
    IF i < iSampleCnt THEN
        fDev := aWeightMg[i] - fMean; // mg − mg = mg / [mg] minus [mg] = [mg]
        fSqSum := fSqSum + (fDev * fDev); // mg × mg = mg² / [mg] × [mg] = [mg^2]
    END_IF
END_FOR
fStd := SQRT(fSqSum / INT_TO_REAL(iSampleCnt - 1)); // mg² ÷ 无量纲 开方 = mg / sqrt([mg^2] / [-]) = [mg]

// 段 5｜RSD 与合格判定
fRsdPct := (fStd / fMean) * 100.0; // mg ÷ mg × 100 = % / [mg] / [mg] × 100 = [%]
IF NOT (fRsdPct > -1.0E30 AND fRsdPct < 1.0E30) THEN
    RETURN; // 结果非有限再拦一次 [-] / second finiteness gate [-]
END_IF
xPass := fRsdPct <= fRsdLimitPct; // 直比上限，禁浮点等值 [-] / direct compare, no float equality [-]
iN := iSampleCnt; // 回填实际样本数 [个] / report the count used [count]
FC_DL_TabletWeightRsdCalc := fRsdPct; // 返回 RSD [%] / return the RSD [%]
END_FUNCTION

(* ---- FC_DL_TankVolumeHoriCyl.st ---- *)
// ==============================================================================
// 组件名 Component  : FC_DL_TankVolumeHoriCyl
// 分类   Category   : DL_Process
// 前缀   Naming     : FC_DL_ ｜ b/f 类型前缀制（R265）
// 版本   Version    : 1.0.0
// 复杂度 Complexity  : 中
// 功能   Purpose    : 卧式圆柱罐液位 - 体积几何解析换算：弦高 → 弓形面积
//                      → 体积（fVol = L * (r²*acos((r-h)/r) − (r−h)*
//                      sqrt(max(0, 2rh − h²)))），h = fLevel 钳位 [0, 2r]；
//                      百分比出口按满罐体积归一。纵坡参数 fTiltDeg 本版
//                      按平面近似支持（> 0 时置 bApprox 提示近似）。
// 文件互引声明 Split : FB_DL_TankLevelStrapping（DL_Process）为查表标定法
//                      （折点表 + 标定核对），本件为几何解析法（公式直算，
//                      零折点依赖），两法勿混用——有标定表用查表件，无表
//                      用本件（R216 双向互引）。
// 开源溯源 Origin    : 道莅原创（弓形面积为公开几何公式，本实现 clean-room，
//                      未复制任何源码行）
// 许可证 License    : MIT
// 参考   Reference  : IEC 61131-3:2013 §6.6.2 函数语义；ACOS / SQRT 为 IEC
//                      标准数学函数；弓形面积公开几何公式（借定义，不抄实现）
// 平台   Platform   : 纯 IEC 61131-3（LREAL 四则 / ACOS / SQRT），三平台通用
// 依赖   Depends    : 无（零委托、零库件；ACOS / SQRT 为 IEC 标准函数）
// 归属 Ownership     : 本件无 TYPE 声明；全部引脚为 IEC 标准原生类型。
// ------------------------------------------------------------------
// 边界 Boundary     :
//   一 组态 / 输入闸（逐项点名，R272）：fDiam <= 0、fLength <= 0、
//      fDiam / fLength / fLevel 任一非有限（NaN 自反判 + Inf 差值自反判 +
//      幅值 1e30 上界）→ bValid = FALSE、双出口归零早退（故障级 303A）；
//   二 液位钳位：h 钳 [0, 2r]（负值钳 0、超高罐顶钳 2r，安全侧归一，
//      信息级 303C 文档语义——本件无 eErr 出口，钳位出口与正常出口
//      同形无独立通道，不另设出口位，R90 反证句）；
//   三 acos 定义域防护：(r - h) / r 钳 [-1, 1]（边界二钳位后 h/r 在
//      [0, 1]，q = 1 - h/r 在 [0, 1]，钳位为防御性双保险，防浮点边缘
//      越域）；除法分母 r > 0 已由组态闸证明；
//   四 被开方数 max(0, 2rh − h²)：h 在 [0, 2r] 已证非负，再叠 max(0,·)
//      双保险，SQRT 入参恒非负；
//   五 百分比分母防零：fVfull = PI*r²*L，由组态闸（fDiam > 0 → r > 0、
//      fLength > 0）证明 fVfull > 0，除法安全（反证句写死）；
//   六 纵坡近似口径：fTiltDeg > 0 → bApprox = TRUE（平面近似，体积按
//      平罐公式给出）；fTiltDeg 非有限 → 同置 bApprox = TRUE 并按 0
//      处理（信息级 303B）；
//   七 结果非有限防御：体积 / 百分比出口算后复检非有限（NaN / Inf /
//      幅值上界），越限即 bValid = FALSE、双出口归零（R273 连续量出口
//      非有限防护）；
//   八 纯函数：无记忆量、无定时器、无边沿实例，每调用重算；
//   九 除法仅两处（h/r 与 fVolM3/fVfull），分母已证非零；无全局、
//      无外部变量、无物理地址。
// 错误码 Codes      :
//   16#0006_303A【故障级】组态 / 输入非法（fDiam / fLength 域非法或任一
//                引脚非有限），bValid = FALSE、双出口归零早退
//   16#0006_303B【信息级】纵坡非零（或非有限按 0 处理），平面近似口径
//                （bApprox = TRUE 通道）
//   16#0006_303C【信息级】液位越界已钳位 [0, 2r]（静默安全侧归一，
//                文档级语义，无独立出口通道）
//   注：本件引脚契约按任务定稿无独立 eErr 出口，故障语义经 bValid /
//   bApprox / 双出口组合表达。
// 验收 Acceptance   :
//   算法已证（脚本）：未跑 ｜ 编译器已证（三平台）：未跑
//   V1 r=1、L=2、h=0 → 体积 0；h=2r → 满罐 PI*r²*L ≈ 6.283 m³、fPct = 100
//   V2 r=1、L=2、h=1（半罐）→ 弓形 = 半圆面积 PI/2 → 体积 ≈ 3.1416、fPct = 50
//   V3 fLevel = -0.5 → 钳 0；fLevel = 5（> 2r）→ 钳 2r
//   V4 fDiam = 0 / 负 → bValid = FALSE；fLevel = NaN → bValid = FALSE
//   V5 fTiltDeg = 3 → bApprox = TRUE（体积仍按平面近似给出）
//   V6 fTiltDeg = NaN → bApprox = TRUE、按 0 处理
// 修订记录 Revision  :
//   2026-11-22  v1.0.0  R65 首版（批 3 · 序号 8）
// ==============================================================================
FUNCTION FC_DL_TankVolumeHoriCyl : BOOL
VAR_INPUT
    fLevel   : LREAL;            // 液位高度 [m]，罐底为 0 / the liquid level, the tank bottom is zero
    fDiam    : LREAL;            // 罐内径 [m]，须 > 0 / the inner diameter, above zero
    fLength  : LREAL;            // 罐筒体长度 [m]，须 > 0 / the shell length, above zero
    fTiltDeg : LREAL := 0.0;     // 纵坡 [deg]，本版平面近似，> 0 置 bApprox / the longitudinal tilt, plane approximation
END_VAR
VAR_OUTPUT
    fVolM3  : LREAL;             // 折算体积 [m³]，无效时 0.0 / the converted volume, zero when invalid
    fPct    : LREAL;             // 体积百分比 [%]，按满罐归一 / the volume percent of the full tank
    bValid  : BOOL;              // 结果可用 [-] / the result usable flag
    bApprox : BOOL;              // 近似口径提示 [-]，纵坡非零 / the approximation flag, a nonzero tilt
END_VAR
VAR
    r         : LREAL;           // 罐半径 [m] / the tank radius
    h         : LREAL;           // 钳位后弦高 [m] / the clamped chord height
    q         : LREAL;           // acos 入参（(r-h)/r）[-] / the acos argument
    fUnder    : LREAL;           // 被开方数 2rh − h² [m²] / the radicand
    fSegArea  : LREAL;           // 弓形截面积 [m²] / the circular segment area
    fVfull    : LREAL;           // 满罐体积 [m³] / the full tank volume
    bTiltBad  : BOOL;            // 纵坡非有限标志 [-] / the tilt fault flag
END_VAR
VAR CONSTANT
    DL_TVC_PI   : LREAL := 3.14159265358979; // 圆周率 [-] / the pi constant
    DL_TVC_FMAX : LREAL := 1.0E30;           // 非有限筛查幅值上限 [m] / the finiteness screening cap
END_VAR

// 段 1｜返回值与全部出口预置（R45 四段式第一段）/ segment 1, the preset of the return and all outlets
FC_DL_TankVolumeHoriCyl := FALSE; // 返回值预置假 / preset the return false
fVolM3  := 0.0;                  // 体积出口预置零 [m³] / preset the volume zero
fPct    := 0.0;                  // 百分比出口预置零 [%] / preset the percent zero
bValid  := FALSE;                // 有效标志预置假 / preset the validity false
bApprox := FALSE;                // 近似提示预置假 / preset the approximation flag false

// 段 2｜组态 / 输入闸（边界一：域 + 非有限逐项点名，R272）/ segment 2, the configuration and input gate
IF (fDiam <= 0.0) OR (fLength <= 0.0)                             // 几何域非法 / an illegal geometry
OR (fLevel <> fLevel) OR ((fLevel - fLevel) <> 0.0) OR (ABS(fLevel) > DL_TVC_FMAX)   // fLevel 非有限 / fLevel non finite
OR (fDiam <> fDiam) OR ((fDiam - fDiam) <> 0.0) OR (ABS(fDiam) > DL_TVC_FMAX)        // fDiam 非有限 / fDiam non finite
OR (fLength <> fLength) OR ((fLength - fLength) <> 0.0) OR (ABS(fLength) > DL_TVC_FMAX) THEN // fLength 非有限 / fLength non finite
    fVolM3 := 0.0;               // 体积归零 [m³] / zero the volume
    fPct   := 0.0;               // 百分比归零 [%] / zero the percent
    bValid := FALSE;             // 故障级 303A：拒绝计算 / refuse the calculation
    RETURN;                      // 早退 / early return
END_IF

// 段 3｜纵坡近似口径（边界六：> 0 置近似，非有限按 0 处理并置近似）/ segment 3, the tilt approximation flag
bTiltBad := (fTiltDeg <> fTiltDeg) OR ((fTiltDeg - fTiltDeg) <> 0.0) OR (ABS(fTiltDeg) > DL_TVC_FMAX); // 纵坡非有限 / the tilt non finite
IF (fTiltDeg > 0.0) OR bTiltBad THEN // 纵坡生效或无效 / the tilt active or invalid
    bApprox := TRUE;             // 信息级 303B：平面近似口径 / the approximation flag raised
END_IF

// 段 4｜半径与液位钳位（边界二：h 钳 [0, 2r]）/ segment 4, the radius and the level clamp
r := fDiam / 2.0;                // 半径 [m]（分母 2.0 为常量，零除面消除）/ the radius, a constant divisor
h := fLevel;                     // 弦高接管 [m] / take the level as the chord height
IF h < 0.0 THEN                  // 液位低于罐底 / the level under the bottom
    h := 0.0;                    // 钳 0（信息级 303C）/ clamp to zero
END_IF
IF h > (2.0 * r) THEN            // 液位超过罐顶 / the level over the top
    h := 2.0 * r;                // 钳 2r（信息级 303C）/ clamp to the full bore
END_IF

// 段 5｜弓形面积解析（边界三 / 四：acos 定义域钳位 + 被开方数非负双保险）/ segment 5, the segment area
q := 1.0 - (h / r);              // acos 入参 (r - h)/r（分母 r > 0 已由组态闸证明）/ the acos argument, the divisor proven above zero
IF q > 1.0 THEN                  // 上越域防御（浮点边缘双保险）/ an upper domain defense
    q := 1.0;                    // 钳回 1.0 / clamp to one
END_IF
IF q < -1.0 THEN                 // 下越域防御 / a lower domain defense
    q := -1.0;                   // 钳回 -1.0 / clamp to minus one
END_IF
fUnder := (2.0 * r * h) - (h * h); // 被开方数 2rh − h² [m²] / the radicand
IF fUnder < 0.0 THEN             // 浮点边缘微负防御（边界四）/ a tiny negative defense
    fUnder := 0.0;               // 钳 0（max(0, ·) 口径）/ clamp to zero
END_IF
fSegArea := (r * r * ACOS(q)) - ((r - h) * SQRT(fUnder)); // 弓形面积公式 [m²] / the segment area formula

// 段 6｜体积与百分比折算（边界五：分母 fVfull > 0 反证已写死）/ segment 6, the volume and the percent
fVolM3 := fLength * fSegArea;    // 体积 = 长度 × 弓形面积 [m³] / the volume as length times the segment area
fVfull := DL_TVC_PI * r * r * fLength; // 满罐体积 [m³]（r > 0 与 L > 0 已证）/ the full volume, proven above zero
fPct   := (fVolM3 / fVfull) * 100.0;   // 百分比 [%]（分母已证非零）/ the percent, the divisor proven

// 段 7｜结果非有限防御（边界七：连续量出口 R273 防护）/ segment 7, the result finiteness defense
IF (fVolM3 <> fVolM3) OR ((fVolM3 - fVolM3) <> 0.0) OR (ABS(fVolM3) > DL_TVC_FMAX) THEN // 体积非有限 / a non finite volume
    fVolM3 := 0.0;               // 体积归零 [m³] / zero the volume
    fPct   := 0.0;               // 百分比归零 [%] / zero the percent
    bValid := FALSE;             // 拒绝输出 / refuse the output
    RETURN;                      // 早退 / early return
END_IF

// 段 8｜统一出口 / segment 8, the unified outlet
bValid := TRUE;                  // 结果可用 / the result usable
FC_DL_TankVolumeHoriCyl := TRUE; // 返回成功 / return success
END_FUNCTION
